(* IEC 61131-3 sources: stf-hw/web/public/sil, 1 file *)

(* ---- stf_plc.st ---- *)
(* STF Upgrade 12 - PLC program, IEC 61131-3 Structured Text. Generated by stf-cad/hbw/sil/iec.py *)
(* from the proven models; compile with MatIEC (iec2c). Task: 5 ms. *)

(* -1 / 0 / +1: which way to drive an axis toward its target; 0 inside the brake lead *)
FUNCTION Drive : INT
VAR_INPUT
    Pos, Tgt, Lead : REAL;
END_VAR
IF Tgt - Pos > Lead THEN Drive := 1; ELSIF Pos - Tgt > Lead THEN Drive := -1; ELSE Drive := 0; END_IF;
END_FUNCTION

(* HBW crane: travel, lift, Ausleger. Generated by stf-cad/hbw/sil/iec.py from the proven motion (control.py); do not edit. *)
FUNCTION_BLOCK FB_Crane
VAR_INPUT
    Enable : BOOL;        (* K0 safety relay OK AND mode = AUTO *)
    Ack : BOOL;           (* HMI acknowledge *)
    Reset : BOOL;         (* S3 reset, via the safety relay *)
    Cmd : INT;            (* job to start (0 = none), taken when READY *)
    Arg1 : INT;           (* binding: slot / bay / slot pair index *)
    I1 : BOOL;           (* reference switch horizontal *)
    I4 : BOOL;           (* reference switch vertical *)
    I5 : BOOL;           (* reference switch cantilever front *)
    I6 : BOOL;           (* reference switch cantilever back *)
    PosTravel : REAL;     (* travel, from the encoder counter *)
    PosLift : REAL;     (* lift, from the encoder counter *)
END_VAR
VAR_OUTPUT
    Q3 : BOOL;           (* horizontal towards rack (M2) *)
    Q4 : BOOL;           (* horizontal towards belt (M2) *)
    Q5 : BOOL;           (* vertical axis down (M3) *)
    Q6 : BOOL;           (* vertical axis up (M3) *)
    Q7 : BOOL;           (* cantilever forward (M4) *)
    Q8 : BOOL;           (* cantilever back (M4) *)
    Ready, Busy, Done, Fault : BOOL;   (* Done: one scan, when a job ends *)
    Alarm : INT;          (* the state whose watchdog tripped *)
    Sn : INT;             (* the active state *)
END_VAR
VAR
    Prev : INT := -1;
    Job, B1 : INT;
    Wd : TON;             (* step watchdog *)
    Tm : TON;             (* step timer *)
    WdTime : TIME;        (* the active state's watchdog; 0 = none *)
END_VAR
VAR CONSTANT
    TG_STORE_RETRIEVE_TRAVEL : ARRAY[1..143, 1..23] OF REAL := [0.0, 0.0, 0.0, 0.0, 0.0, 0.0, 0.0, 0.0, 0.0, 0.0, 0.0, 0.0, 0.0, 0.0, 0.0, 0.0, 0.0, 0.0, 0.0, 0.0, 0.0, 0.0, 0.0, 0.0, 0.0, 0.0, 0.0, 0.0, 120.0, 0.0, 0.0, 0.0, 0.0, 0.0, 240.0, 0.0, 0.0, 0.0, 0.0, 0.0, 665.0, 0.0, 0.0, 0.0, 0.0, 0.0, 0.0, 0.0, 0.0, 0.0, 0.0, 120.0, 0.0, 0.0, 0.0, 0.0, 0.0, 360.0, 0.0, 0.0, 0.0, 0.0, 0.0, 665.0, 0.0, 0.0, 0.0, 0.0, 0.0, 0.0, 0.0, 0.0, 0.0, 0.0, 120.0, 0.0, 0.0, 0.0, 0.0, 0.0, 480.0, 0.0, 0.0, 0.0, 0.0, 0.0, 665.0, 0.0, 0.0, 0.0, 0.0, 0.0, 0.0, 0.0, 0.0, 0.0, 0.0, 120.0, 0.0, 0.0, 0.0, 0.0, 0.0, 120.0, 0.0, 0.0, 0.0, 0.0, 0.0, 665.0, 0.0, 0.0, 0.0, 0.0, 0.0, 0.0, 0.0, 0.0, 0.0, 0.0, 120.0, 0.0, 0.0, 0.0, 0.0, 0.0, 240.0, 0.0, 0.0, 0.0, 0.0, 0.0, 665.0, 0.0, 0.0, 0.0, 0.0, 0.0, 0.0, 0.0, 0.0, 0.0, 0.0, 120.0, 0.0, 0.0, 0.0, 0.0, 0.0, 360.0, 0.0, 0.0, 0.0, 0.0, 0.0, 665.0, 0.0, 0.0, 0.0, 0.0, 0.0, 0.0, 0.0, 0.0, 0.0, 0.0, 120.0, 0.0, 0.0, 0.0, 0.0, 0.0, 480.0, 0.0, 0.0, 0.0, 0.0, 0.0, 665.0, 0.0, 0.0, 0.0, 0.0, 0.0, 0.0, 0.0, 0.0, 0.0, 0.0, 120.0, 0.0, 0.0, 0.0, 0.0, 0.0, 120.0, 0.0, 0.0, 0.0, 0.0, 0.0, 665.0, 0.0, 0.0, 0.0, 0.0, 0.0, 0.0, 0.0, 0.0, 0.0, 0.0, 120.0, 0.0, 0.0, 0.0, 0.0, 0.0, 240.0, 0.0, 0.0, 0.0, 0.0, 0.0, 665.0, 0.0, 0.0, 0.0, 0.0, 0.0, 0.0, 0.0, 0.0, 0.0, 0.0, 120.0, 0.0, 0.0, 0.0, 0.0, 0.0, 360.0, 0.0, 0.0, 0.0, 0.0, 0.0, 665.0, 0.0, 0.0, 0.0, 0.0, 0.0, 0.0, 0.0, 0.0, 0.0, 0.0, 120.0, 0.0, 0.0, 0.0, 0.0, 0.0, 480.0, 0.0, 0.0, 0.0, 0.0, 0.0, 665.0, 0.0, 0.0, 0.0, 0.0, 0.0, 0.0, 0.0, 0.0, 0.0, 0.0, 240.0, 0.0, 0.0, 0.0, 0.0, 0.0, 120.0, 0.0, 0.0, 0.0, 0.0, 0.0, 665.0, 0.0, 0.0, 0.0, 0.0, 0.0, 0.0, 0.0, 0.0, 0.0, 0.0, 0.0, 0.0, 0.0, 0.0, 0.0, 0.0, 0.0, 0.0, 0.0, 0.0, 0.0, 0.0, 0.0, 0.0, 0.0, 0.0, 0.0, 0.0, 0.0, 0.0, 0.0, 0.0, 0.0, 240.0, 0.0, 0.0, 0.0, 0.0, 0.0, 360.0, 0.0, 0.0, 0.0, 0.0, 0.0, 665.0, 0.0, 0.0, 0.0, 0.0, 0.0, 0.0, 0.0, 0.0, 0.0, 0.0, 240.0, 0.0, 0.0, 0.0, 0.0, 0.0, 480.0, 0.0, 0.0, 0.0, 0.0, 0.0, 665.0, 0.0, 0.0, 0.0, 0.0, 0.0, 0.0, 0.0, 0.0, 0.0, 0.0, 240.0, 0.0, 0.0, 0.0, 0.0, 0.0, 120.0, 0.0, 0.0, 0.0, 0.0, 0.0, 665.0, 0.0, 0.0, 0.0, 0.0, 0.0, 0.0, 0.0, 0.0, 0.0, 0.0, 240.0, 0.0, 0.0, 0.0, 0.0, 0.0, 240.0, 0.0, 0.0, 0.0, 0.0, 0.0, 665.0, 0.0, 0.0, 0.0, 0.0, 0.0, 0.0, 0.0, 0.0, 0.0, 0.0, 240.0, 0.0, 0.0, 0.0, 0.0, 0.0, 360.0, 0.0, 0.0, 0.0, 0.0, 0.0, 665.0, 0.0, 0.0, 0.0, 0.0, 0.0, 0.0, 0.0, 0.0, 0.0, 0.0, 240.0, 0.0, 0.0, 0.0, 0.0, 0.0, 480.0, 0.0, 0.0, 0.0, 0.0, 0.0, 665.0, 0.0, 0.0, 0.0, 0.0, 0.0, 0.0, 0.0, 0.0, 0.0, 0.0, 240.0, 0.0, 0.0, 0.0, 0.0, 0.0, 120.0, 0.0, 0.0, 0.0, 0.0, 0.0, 665.0, 0.0, 0.0, 0.0, 0.0, 0.0, 0.0, 0.0, 0.0, 0.0, 0.0, 240.0, 0.0, 0.0, 0.0, 0.0, 0.0, 240.0, 0.0, 0.0, 0.0, 0.0, 0.0, 665.0, 0.0, 0.0, 0.0, 0.0, 0.0, 0.0, 0.0, 0.0, 0.0, 0.0, 240.0, 0.0, 0.0, 0.0, 0.0, 0.0, 360.0, 0.0, 0.0, 0.0, 0.0, 0.0, 665.0, 0.0, 0.0, 0.0, 0.0, 0.0, 0.0, 0.0, 0.0, 0.0, 0.0, 240.0, 0.0, 0.0, 0.0, 0.0, 0.0, 480.0, 0.0, 0.0, 0.0, 0.0, 0.0, 665.0, 0.0, 0.0, 0.0, 0.0, 0.0, 0.0, 0.0, 0.0, 0.0, 0.0, 360.0, 0.0, 0.0, 0.0, 0.0, 0.0, 120.0, 0.0, 0.0, 0.0, 0.0, 0.0, 665.0, 0.0, 0.0, 0.0, 0.0, 0.0, 0.0, 0.0, 0.0, 0.0, 0.0, 360.0, 0.0, 0.0, 0.0, 0.0, 0.0, 240.0, 0.0, 0.0, 0.0, 0.0, 0.0, 665.0, 0.0, 0.0, 0.0, 0.0, 0.0, 0.0, 0.0, 0.0, 0.0, 0.0, 0.0, 0.0, 0.0, 0.0, 0.0, 0.0, 0.0, 0.0, 0.0, 0.0, 0.0, 0.0, 0.0, 0.0, 0.0, 0.0, 0.0, 0.0, 0.0, 0.0, 0.0, 0.0, 0.0, 360.0, 0.0, 0.0, 0.0, 0.0, 0.0, 480.0, 0.0, 0.0, 0.0, 0.0, 0.0, 665.0, 0.0, 0.0, 0.0, 0.0, 0.0, 0.0, 0.0, 0.0, 0.0, 0.0, 360.0, 0.0, 0.0, 0.0, 0.0, 0.0, 120.0, 0.0, 0.0, 0.0, 0.0, 0.0, 665.0, 0.0, 0.0, 0.0, 0.0, 0.0, 0.0, 0.0, 0.0, 0.0, 0.0, 360.0, 0.0, 0.0, 0.0, 0.0, 0.0, 240.0, 0.0, 0.0, 0.0, 0.0, 0.0, 665.0, 0.0, 0.0, 0.0, 0.0, 0.0, 0.0, 0.0, 0.0, 0.0, 0.0, 360.0, 0.0, 0.0, 0.0, 0.0, 0.0, 360.0, 0.0, 0.0, 0.0, 0.0, 0.0, 665.0, 0.0, 0.0, 0.0, 0.0, 0.0, 0.0, 0.0, 0.0, 0.0, 0.0, 360.0, 0.0, 0.0, 0.0, 0.0, 0.0, 480.0, 0.0, 0.0, 0.0, 0.0, 0.0, 665.0, 0.0, 0.0, 0.0, 0.0, 0.0, 0.0, 0.0, 0.0, 0.0, 0.0, 360.0, 0.0, 0.0, 0.0, 0.0, 0.0, 120.0, 0.0, 0.0, 0.0, 0.0, 0.0, 665.0, 0.0, 0.0, 0.0, 0.0, 0.0, 0.0, 0.0, 0.0, 0.0, 0.0, 360.0, 0.0, 0.0, 0.0, 0.0, 0.0, 240.0, 0.0, 0.0, 0.0, 0.0, 0.0, 665.0, 0.0, 0.0, 0.0, 0.0, 0.0, 0.0, 0.0, 0.0, 0.0, 0.0, 360.0, 0.0, 0.0, 0.0, 0.0, 0.0, 360.0, 0.0, 0.0, 0.0, 0.0, 0.0, 665.0, 0.0, 0.0, 0.0, 0.0, 0.0, 0.0, 0.0, 0.0, 0.0, 0.0, 360.0, 0.0, 0.0, 0.0, 0.0, 0.0, 480.0, 0.0, 0.0, 0.0, 0.0, 0.0, 665.0, 0.0, 0.0, 0.0, 0.0, 0.0, 0.0, 0.0, 0.0, 0.0, 0.0, 480.0, 0.0, 0.0, 0.0, 0.0, 0.0, 120.0, 0.0, 0.0, 0.0, 0.0, 0.0, 665.0, 0.0, 0.0, 0.0, 0.0, 0.0, 0.0, 0.0, 0.0, 0.0, 0.0, 480.0, 0.0, 0.0, 0.0, 0.0, 0.0, 240.0, 0.0, 0.0, 0.0, 0.0, 0.0, 665.0, 0.0, 0.0, 0.0, 0.0, 0.0, 0.0, 0.0, 0.0, 0.0, 0.0, 480.0, 0.0, 0.0, 0.0, 0.0, 0.0, 360.0, 0.0, 0.0, 0.0, 0.0, 0.0, 665.0, 0.0, 0.0, 0.0, 0.0, 0.0, 0.0, 0.0, 0.0, 0.0, 0.0, 0.0, 0.0, 0.0, 0.0, 0.0, 0.0, 0.0, 0.0, 0.0, 0.0, 0.0, 0.0, 0.0, 0.0, 0.0, 0.0, 0.0, 0.0, 0.0, 0.0, 0.0, 0.0, 0.0, 480.0, 0.0, 0.0, 0.0, 0.0, 0.0, 120.0, 0.0, 0.0, 0.0, 0.0, 0.0, 665.0, 0.0, 0.0, 0.0, 0.0, 0.0, 0.0, 0.0, 0.0, 0.0, 0.0, 480.0, 0.0, 0.0, 0.0, 0.0, 0.0, 240.0, 0.0, 0.0, 0.0, 0.0, 0.0, 665.0, 0.0, 0.0, 0.0, 0.0, 0.0, 0.0, 0.0, 0.0, 0.0, 0.0, 480.0, 0.0, 0.0, 0.0, 0.0, 0.0, 360.0, 0.0, 0.0, 0.0, 0.0, 0.0, 665.0, 0.0, 0.0, 0.0, 0.0, 0.0, 0.0, 0.0, 0.0, 0.0, 0.0, 480.0, 0.0, 0.0, 0.0, 0.0, 0.0, 480.0, 0.0, 0.0, 0.0, 0.0, 0.0, 665.0, 0.0, 0.0, 0.0, 0.0, 0.0, 0.0, 0.0, 0.0, 0.0, 0.0, 480.0, 0.0, 0.0, 0.0, 0.0, 0.0, 120.0, 0.0, 0.0, 0.0, 0.0, 0.0, 665.0, 0.0, 0.0, 0.0, 0.0, 0.0, 0.0, 0.0, 0.0, 0.0, 0.0, 480.0, 0.0, 0.0, 0.0, 0.0, 0.0, 240.0, 0.0, 0.0, 0.0, 0.0, 0.0, 665.0, 0.0, 0.0, 0.0, 0.0, 0.0, 0.0, 0.0, 0.0, 0.0, 0.0, 480.0, 0.0, 0.0, 0.0, 0.0, 0.0, 360.0, 0.0, 0.0, 0.0, 0.0, 0.0, 665.0, 0.0, 0.0, 0.0, 0.0, 0.0, 0.0, 0.0, 0.0, 0.0, 0.0, 480.0, 0.0, 0.0, 0.0, 0.0, 0.0, 480.0, 0.0, 0.0, 0.0, 0.0, 0.0, 665.0, 0.0, 0.0, 0.0, 0.0, 0.0, 0.0, 0.0, 0.0, 0.0, 0.0, 120.0, 0.0, 0.0, 0.0, 0.0, 0.0, 120.0, 0.0, 0.0, 0.0, 0.0, 0.0, 665.0, 0.0, 0.0, 0.0, 0.0, 0.0, 0.0, 0.0, 0.0, 0.0, 0.0, 120.0, 0.0, 0.0, 0.0, 0.0, 0.0, 240.0, 0.0, 0.0, 0.0, 0.0, 0.0, 665.0, 0.0, 0.0, 0.0, 0.0, 0.0, 0.0, 0.0, 0.0, 0.0, 0.0, 120.0, 0.0, 0.0, 0.0, 0.0, 0.0, 360.0, 0.0, 0.0, 0.0, 0.0, 0.0, 665.0, 0.0, 0.0, 0.0, 0.0, 0.0, 0.0, 0.0, 0.0, 0.0, 0.0, 120.0, 0.0, 0.0, 0.0, 0.0, 0.0, 480.0, 0.0, 0.0, 0.0, 0.0, 0.0, 665.0, 0.0, 0.0, 0.0, 0.0, 0.0, 0.0, 0.0, 0.0, 0.0, 0.0, 0.0, 0.0, 0.0, 0.0, 0.0, 0.0, 0.0, 0.0, 0.0, 0.0, 0.0, 0.0, 0.0, 0.0, 0.0, 0.0, 0.0, 0.0, 0.0, 0.0, 0.0, 0.0, 0.0, 120.0, 0.0, 0.0, 0.0, 0.0, 0.0, 240.0, 0.0, 0.0, 0.0, 0.0, 0.0, 665.0, 0.0, 0.0, 0.0, 0.0, 0.0, 0.0, 0.0, 0.0, 0.0, 0.0, 120.0, 0.0, 0.0, 0.0, 0.0, 0.0, 360.0, 0.0, 0.0, 0.0, 0.0, 0.0, 665.0, 0.0, 0.0, 0.0, 0.0, 0.0, 0.0, 0.0, 0.0, 0.0, 0.0, 120.0, 0.0, 0.0, 0.0, 0.0, 0.0, 480.0, 0.0, 0.0, 0.0, 0.0, 0.0, 665.0, 0.0, 0.0, 0.0, 0.0, 0.0, 0.0, 0.0, 0.0, 0.0, 0.0, 120.0, 0.0, 0.0, 0.0, 0.0, 0.0, 120.0, 0.0, 0.0, 0.0, 0.0, 0.0, 665.0, 0.0, 0.0, 0.0, 0.0, 0.0, 0.0, 0.0, 0.0, 0.0, 0.0, 120.0, 0.0, 0.0, 0.0, 0.0, 0.0, 240.0, 0.0, 0.0, 0.0, 0.0, 0.0, 665.0, 0.0, 0.0, 0.0, 0.0, 0.0, 0.0, 0.0, 0.0, 0.0, 0.0, 120.0, 0.0, 0.0, 0.0, 0.0, 0.0, 360.0, 0.0, 0.0, 0.0, 0.0, 0.0, 665.0, 0.0, 0.0, 0.0, 0.0, 0.0, 0.0, 0.0, 0.0, 0.0, 0.0, 120.0, 0.0, 0.0, 0.0, 0.0, 0.0, 480.0, 0.0, 0.0, 0.0, 0.0, 0.0, 665.0, 0.0, 0.0, 0.0, 0.0, 0.0, 0.0, 0.0, 0.0, 0.0, 0.0, 240.0, 0.0, 0.0, 0.0, 0.0, 0.0, 120.0, 0.0, 0.0, 0.0, 0.0, 0.0, 665.0, 0.0, 0.0, 0.0, 0.0, 0.0, 0.0, 0.0, 0.0, 0.0, 0.0, 240.0, 0.0, 0.0, 0.0, 0.0, 0.0, 240.0, 0.0, 0.0, 0.0, 0.0, 0.0, 665.0, 0.0, 0.0, 0.0, 0.0, 0.0, 0.0, 0.0, 0.0, 0.0, 0.0, 240.0, 0.0, 0.0, 0.0, 0.0, 0.0, 360.0, 0.0, 0.0, 0.0, 0.0, 0.0, 665.0, 0.0, 0.0, 0.0, 0.0, 0.0, 0.0, 0.0, 0.0, 0.0, 0.0, 240.0, 0.0, 0.0, 0.0, 0.0, 0.0, 480.0, 0.0, 0.0, 0.0, 0.0, 0.0, 665.0, 0.0, 0.0, 0.0, 0.0, 0.0, 0.0, 0.0, 0.0, 0.0, 0.0, 240.0, 0.0, 0.0, 0.0, 0.0, 0.0, 120.0, 0.0, 0.0, 0.0, 0.0, 0.0, 665.0, 0.0, 0.0, 0.0, 0.0, 0.0, 0.0, 0.0, 0.0, 0.0, 0.0, 0.0, 0.0, 0.0, 0.0, 0.0, 0.0, 0.0, 0.0, 0.0, 0.0, 0.0, 0.0, 0.0, 0.0, 0.0, 0.0, 0.0, 0.0, 0.0, 0.0, 0.0, 0.0, 0.0, 240.0, 0.0, 0.0, 0.0, 0.0, 0.0, 360.0, 0.0, 0.0, 0.0, 0.0, 0.0, 665.0, 0.0, 0.0, 0.0, 0.0, 0.0, 0.0, 0.0, 0.0, 0.0, 0.0, 240.0, 0.0, 0.0, 0.0, 0.0, 0.0, 480.0, 0.0, 0.0, 0.0, 0.0, 0.0, 665.0, 0.0, 0.0, 0.0, 0.0, 0.0, 0.0, 0.0, 0.0, 0.0, 0.0, 240.0, 0.0, 0.0, 0.0, 0.0, 0.0, 120.0, 0.0, 0.0, 0.0, 0.0, 0.0, 665.0, 0.0, 0.0, 0.0, 0.0, 0.0, 0.0, 0.0, 0.0, 0.0, 0.0, 240.0, 0.0, 0.0, 0.0, 0.0, 0.0, 240.0, 0.0, 0.0, 0.0, 0.0, 0.0, 665.0, 0.0, 0.0, 0.0, 0.0, 0.0, 0.0, 0.0, 0.0, 0.0, 0.0, 240.0, 0.0, 0.0, 0.0, 0.0, 0.0, 360.0, 0.0, 0.0, 0.0, 0.0, 0.0, 665.0, 0.0, 0.0, 0.0, 0.0, 0.0, 0.0, 0.0, 0.0, 0.0, 0.0, 240.0, 0.0, 0.0, 0.0, 0.0, 0.0, 480.0, 0.0, 0.0, 0.0, 0.0, 0.0, 665.0, 0.0, 0.0, 0.0, 0.0, 0.0, 0.0, 0.0, 0.0, 0.0, 0.0, 360.0, 0.0, 0.0, 0.0, 0.0, 0.0, 120.0, 0.0, 0.0, 0.0, 0.0, 0.0, 665.0, 0.0, 0.0, 0.0, 0.0, 0.0, 0.0, 0.0, 0.0, 0.0, 0.0, 360.0, 0.0, 0.0, 0.0, 0.0, 0.0, 240.0, 0.0, 0.0, 0.0, 0.0, 0.0, 665.0, 0.0, 0.0, 0.0, 0.0, 0.0, 0.0, 0.0, 0.0, 0.0, 0.0, 360.0, 0.0, 0.0, 0.0, 0.0, 0.0, 360.0, 0.0, 0.0, 0.0, 0.0, 0.0, 665.0, 0.0, 0.0, 0.0, 0.0, 0.0, 0.0, 0.0, 0.0, 0.0, 0.0, 360.0, 0.0, 0.0, 0.0, 0.0, 0.0, 480.0, 0.0, 0.0, 0.0, 0.0, 0.0, 665.0, 0.0, 0.0, 0.0, 0.0, 0.0, 0.0, 0.0, 0.0, 0.0, 0.0, 360.0, 0.0, 0.0, 0.0, 0.0, 0.0, 120.0, 0.0, 0.0, 0.0, 0.0, 0.0, 665.0, 0.0, 0.0, 0.0, 0.0, 0.0, 0.0, 0.0, 0.0, 0.0, 0.0, 360.0, 0.0, 0.0, 0.0, 0.0, 0.0, 240.0, 0.0, 0.0, 0.0, 0.0, 0.0, 665.0, 0.0, 0.0, 0.0, 0.0, 0.0, 0.0, 0.0, 0.0, 0.0, 0.0, 0.0, 0.0, 0.0, 0.0, 0.0, 0.0, 0.0, 0.0, 0.0, 0.0, 0.0, 0.0, 0.0, 0.0, 0.0, 0.0, 0.0, 0.0, 0.0, 0.0, 0.0, 0.0, 0.0, 360.0, 0.0, 0.0, 0.0, 0.0, 0.0, 480.0, 0.0, 0.0, 0.0, 0.0, 0.0, 665.0, 0.0, 0.0, 0.0, 0.0, 0.0, 0.0, 0.0, 0.0, 0.0, 0.0, 360.0, 0.0, 0.0, 0.0, 0.0, 0.0, 120.0, 0.0, 0.0, 0.0, 0.0, 0.0, 665.0, 0.0, 0.0, 0.0, 0.0, 0.0, 0.0, 0.0, 0.0, 0.0, 0.0, 360.0, 0.0, 0.0, 0.0, 0.0, 0.0, 240.0, 0.0, 0.0, 0.0, 0.0, 0.0, 665.0, 0.0, 0.0, 0.0, 0.0, 0.0, 0.0, 0.0, 0.0, 0.0, 0.0, 360.0, 0.0, 0.0, 0.0, 0.0, 0.0, 360.0, 0.0, 0.0, 0.0, 0.0, 0.0, 665.0, 0.0, 0.0, 0.0, 0.0, 0.0, 0.0, 0.0, 0.0, 0.0, 0.0, 360.0, 0.0, 0.0, 0.0, 0.0, 0.0, 480.0, 0.0, 0.0, 0.0, 0.0, 0.0, 665.0, 0.0, 0.0, 0.0, 0.0, 0.0, 0.0, 0.0, 0.0, 0.0, 0.0, 480.0, 0.0, 0.0, 0.0, 0.0, 0.0, 120.0, 0.0, 0.0, 0.0, 0.0, 0.0, 665.0, 0.0, 0.0, 0.0, 0.0, 0.0, 0.0, 0.0, 0.0, 0.0, 0.0, 480.0, 0.0, 0.0, 0.0, 0.0, 0.0, 240.0, 0.0, 0.0, 0.0, 0.0, 0.0, 665.0, 0.0, 0.0, 0.0, 0.0, 0.0, 0.0, 0.0, 0.0, 0.0, 0.0, 480.0, 0.0, 0.0, 0.0, 0.0, 0.0, 360.0, 0.0, 0.0, 0.0, 0.0, 0.0, 665.0, 0.0, 0.0, 0.0, 0.0, 0.0, 0.0, 0.0, 0.0, 0.0, 0.0, 480.0, 0.0, 0.0, 0.0, 0.0, 0.0, 480.0, 0.0, 0.0, 0.0, 0.0, 0.0, 665.0, 0.0, 0.0, 0.0, 0.0, 0.0, 0.0, 0.0, 0.0, 0.0, 0.0, 480.0, 0.0, 0.0, 0.0, 0.0, 0.0, 120.0, 0.0, 0.0, 0.0, 0.0, 0.0, 665.0, 0.0, 0.0, 0.0, 0.0, 0.0, 0.0, 0.0, 0.0, 0.0, 0.0, 480.0, 0.0, 0.0, 0.0, 0.0, 0.0, 240.0, 0.0, 0.0, 0.0, 0.0, 0.0, 665.0, 0.0, 0.0, 0.0, 0.0, 0.0, 0.0, 0.0, 0.0, 0.0, 0.0, 480.0, 0.0, 0.0, 0.0, 0.0, 0.0, 360.0, 0.0, 0.0, 0.0, 0.0, 0.0, 665.0, 0.0, 0.0, 0.0, 0.0, 0.0, 0.0, 0.0, 0.0, 0.0, 0.0, 0.0, 0.0, 0.0, 0.0, 0.0, 0.0, 0.0, 0.0, 0.0, 0.0, 0.0, 0.0, 0.0, 0.0, 0.0, 0.0, 0.0, 0.0, 0.0, 0.0, 0.0, 0.0, 0.0, 480.0, 0.0, 0.0, 0.0, 0.0, 0.0, 120.0, 0.0, 0.0, 0.0, 0.0, 0.0, 665.0, 0.0, 0.0, 0.0, 0.0, 0.0, 0.0, 0.0, 0.0, 0.0, 0.0, 480.0, 0.0, 0.0, 0.0, 0.0, 0.0, 240.0, 0.0, 0.0, 0.0, 0.0, 0.0, 665.0, 0.0, 0.0, 0.0, 0.0, 0.0, 0.0, 0.0, 0.0, 0.0, 0.0, 480.0, 0.0, 0.0, 0.0, 0.0, 0.0, 360.0, 0.0, 0.0, 0.0, 0.0, 0.0, 665.0, 0.0, 0.0, 0.0, 0.0, 0.0, 0.0, 0.0, 0.0, 0.0, 0.0, 480.0, 0.0, 0.0, 0.0, 0.0, 0.0, 480.0, 0.0, 0.0, 0.0, 0.0, 0.0, 665.0, 0.0, 0.0, 0.0, 0.0, 0.0, 0.0, 0.0, 0.0, 0.0, 0.0, 120.0, 0.0, 0.0, 0.0, 0.0, 0.0, 120.0, 0.0, 0.0, 0.0, 0.0, 0.0, 665.0, 0.0, 0.0, 0.0, 0.0, 0.0, 0.0, 0.0, 0.0, 0.0, 0.0, 120.0, 0.0, 0.0, 0.0, 0.0, 0.0, 240.0, 0.0, 0.0, 0.0, 0.0, 0.0, 665.0, 0.0, 0.0, 0.0, 0.0, 0.0, 0.0, 0.0, 0.0, 0.0, 0.0, 120.0, 0.0, 0.0, 0.0, 0.0, 0.0, 360.0, 0.0, 0.0, 0.0, 0.0, 0.0, 665.0, 0.0, 0.0, 0.0, 0.0, 0.0, 0.0, 0.0, 0.0, 0.0, 0.0, 120.0, 0.0, 0.0, 0.0, 0.0, 0.0, 480.0, 0.0, 0.0, 0.0, 0.0, 0.0, 665.0, 0.0, 0.0, 0.0, 0.0, 0.0, 0.0, 0.0, 0.0, 0.0, 0.0, 120.0, 0.0, 0.0, 0.0, 0.0, 0.0, 120.0, 0.0, 0.0, 0.0, 0.0, 0.0, 665.0, 0.0, 0.0, 0.0, 0.0, 0.0, 0.0, 0.0, 0.0, 0.0, 0.0, 120.0, 0.0, 0.0, 0.0, 0.0, 0.0, 240.0, 0.0, 0.0, 0.0, 0.0, 0.0, 665.0, 0.0, 0.0, 0.0, 0.0, 0.0, 0.0, 0.0, 0.0, 0.0, 0.0, 120.0, 0.0, 0.0, 0.0, 0.0, 0.0, 360.0, 0.0, 0.0, 0.0, 0.0, 0.0, 665.0, 0.0, 0.0, 0.0, 0.0, 0.0, 0.0, 0.0, 0.0, 0.0, 0.0, 120.0, 0.0, 0.0, 0.0, 0.0, 0.0, 480.0, 0.0, 0.0, 0.0, 0.0, 0.0, 665.0, 0.0, 0.0, 0.0, 0.0, 0.0, 0.0, 0.0, 0.0, 0.0, 0.0, 0.0, 0.0, 0.0, 0.0, 0.0, 0.0, 0.0, 0.0, 0.0, 0.0, 0.0, 0.0, 0.0, 0.0, 0.0, 0.0, 0.0, 0.0, 0.0, 0.0, 0.0, 0.0, 0.0, 120.0, 0.0, 0.0, 0.0, 0.0, 0.0, 240.0, 0.0, 0.0, 0.0, 0.0, 0.0, 665.0, 0.0, 0.0, 0.0, 0.0, 0.0, 0.0, 0.0, 0.0, 0.0, 0.0, 120.0, 0.0, 0.0, 0.0, 0.0, 0.0, 360.0, 0.0, 0.0, 0.0, 0.0, 0.0, 665.0, 0.0, 0.0, 0.0, 0.0, 0.0, 0.0, 0.0, 0.0, 0.0, 0.0, 120.0, 0.0, 0.0, 0.0, 0.0, 0.0, 480.0, 0.0, 0.0, 0.0, 0.0, 0.0, 665.0, 0.0, 0.0, 0.0, 0.0, 0.0, 0.0, 0.0, 0.0, 0.0, 0.0, 240.0, 0.0, 0.0, 0.0, 0.0, 0.0, 120.0, 0.0, 0.0, 0.0, 0.0, 0.0, 665.0, 0.0, 0.0, 0.0, 0.0, 0.0, 0.0, 0.0, 0.0, 0.0, 0.0, 240.0, 0.0, 0.0, 0.0, 0.0, 0.0, 240.0, 0.0, 0.0, 0.0, 0.0, 0.0, 665.0, 0.0, 0.0, 0.0, 0.0, 0.0, 0.0, 0.0, 0.0, 0.0, 0.0, 240.0, 0.0, 0.0, 0.0, 0.0, 0.0, 360.0, 0.0, 0.0, 0.0, 0.0, 0.0, 665.0, 0.0, 0.0, 0.0, 0.0, 0.0, 0.0, 0.0, 0.0, 0.0, 0.0, 240.0, 0.0, 0.0, 0.0, 0.0, 0.0, 480.0, 0.0, 0.0, 0.0, 0.0, 0.0, 665.0, 0.0, 0.0, 0.0, 0.0, 0.0, 0.0, 0.0, 0.0, 0.0, 0.0, 240.0, 0.0, 0.0, 0.0, 0.0, 0.0, 120.0, 0.0, 0.0, 0.0, 0.0, 0.0, 665.0, 0.0, 0.0, 0.0, 0.0, 0.0, 0.0, 0.0, 0.0, 0.0, 0.0, 240.0, 0.0, 0.0, 0.0, 0.0, 0.0, 240.0, 0.0, 0.0, 0.0, 0.0, 0.0, 665.0, 0.0, 0.0, 0.0, 0.0, 0.0, 0.0, 0.0, 0.0, 0.0, 0.0, 240.0, 0.0, 0.0, 0.0, 0.0, 0.0, 360.0, 0.0, 0.0, 0.0, 0.0, 0.0, 665.0, 0.0, 0.0, 0.0, 0.0, 0.0, 0.0, 0.0, 0.0, 0.0, 0.0, 240.0, 0.0, 0.0, 0.0, 0.0, 0.0, 480.0, 0.0, 0.0, 0.0, 0.0, 0.0, 665.0, 0.0, 0.0, 0.0, 0.0, 0.0, 0.0, 0.0, 0.0, 0.0, 0.0, 240.0, 0.0, 0.0, 0.0, 0.0, 0.0, 120.0, 0.0, 0.0, 0.0, 0.0, 0.0, 665.0, 0.0, 0.0, 0.0, 0.0, 0.0, 0.0, 0.0, 0.0, 0.0, 0.0, 0.0, 0.0, 0.0, 0.0, 0.0, 0.0, 0.0, 0.0, 0.0, 0.0, 0.0, 0.0, 0.0, 0.0, 0.0, 0.0, 0.0, 0.0, 0.0, 0.0, 0.0, 0.0, 0.0, 240.0, 0.0, 0.0, 0.0, 0.0, 0.0, 360.0, 0.0, 0.0, 0.0, 0.0, 0.0, 665.0, 0.0, 0.0, 0.0, 0.0, 0.0, 0.0, 0.0, 0.0, 0.0, 0.0, 240.0, 0.0, 0.0, 0.0, 0.0, 0.0, 480.0, 0.0, 0.0, 0.0, 0.0, 0.0, 665.0, 0.0, 0.0, 0.0, 0.0, 0.0, 0.0, 0.0, 0.0, 0.0, 0.0, 360.0, 0.0, 0.0, 0.0, 0.0, 0.0, 120.0, 0.0, 0.0, 0.0, 0.0, 0.0, 665.0, 0.0, 0.0, 0.0, 0.0, 0.0, 0.0, 0.0, 0.0, 0.0, 0.0, 360.0, 0.0, 0.0, 0.0, 0.0, 0.0, 240.0, 0.0, 0.0, 0.0, 0.0, 0.0, 665.0, 0.0, 0.0, 0.0, 0.0, 0.0, 0.0, 0.0, 0.0, 0.0, 0.0, 360.0, 0.0, 0.0, 0.0, 0.0, 0.0, 360.0, 0.0, 0.0, 0.0, 0.0, 0.0, 665.0, 0.0, 0.0, 0.0, 0.0, 0.0, 0.0, 0.0, 0.0, 0.0, 0.0, 360.0, 0.0, 0.0, 0.0, 0.0, 0.0, 480.0, 0.0, 0.0, 0.0, 0.0, 0.0, 665.0, 0.0, 0.0, 0.0, 0.0, 0.0, 0.0, 0.0, 0.0, 0.0, 0.0, 360.0, 0.0, 0.0, 0.0, 0.0, 0.0, 120.0, 0.0, 0.0, 0.0, 0.0, 0.0, 665.0, 0.0, 0.0, 0.0, 0.0, 0.0, 0.0, 0.0, 0.0, 0.0, 0.0, 360.0, 0.0, 0.0, 0.0, 0.0, 0.0, 240.0, 0.0, 0.0, 0.0, 0.0, 0.0, 665.0, 0.0, 0.0, 0.0, 0.0, 0.0, 0.0, 0.0, 0.0, 0.0, 0.0, 360.0, 0.0, 0.0, 0.0, 0.0, 0.0, 360.0, 0.0, 0.0, 0.0, 0.0, 0.0, 665.0, 0.0, 0.0, 0.0, 0.0, 0.0, 0.0, 0.0, 0.0, 0.0, 0.0, 360.0, 0.0, 0.0, 0.0, 0.0, 0.0, 480.0, 0.0, 0.0, 0.0, 0.0, 0.0, 665.0, 0.0, 0.0, 0.0, 0.0, 0.0, 0.0, 0.0, 0.0, 0.0, 0.0, 360.0, 0.0, 0.0, 0.0, 0.0, 0.0, 120.0, 0.0, 0.0, 0.0, 0.0, 0.0, 665.0, 0.0, 0.0, 0.0, 0.0, 0.0, 0.0, 0.0, 0.0, 0.0, 0.0, 360.0, 0.0, 0.0, 0.0, 0.0, 0.0, 240.0, 0.0, 0.0, 0.0, 0.0, 0.0, 665.0, 0.0, 0.0, 0.0, 0.0, 0.0, 0.0, 0.0, 0.0, 0.0, 0.0, 0.0, 0.0, 0.0, 0.0, 0.0, 0.0, 0.0, 0.0, 0.0, 0.0, 0.0, 0.0, 0.0, 0.0, 0.0, 0.0, 0.0, 0.0, 0.0, 0.0, 0.0, 0.0, 0.0, 360.0, 0.0, 0.0, 0.0, 0.0, 0.0, 480.0, 0.0, 0.0, 0.0, 0.0, 0.0, 665.0, 0.0, 0.0, 0.0, 0.0, 0.0, 0.0, 0.0, 0.0, 0.0, 0.0, 480.0, 0.0, 0.0, 0.0, 0.0, 0.0, 120.0, 0.0, 0.0, 0.0, 0.0, 0.0, 665.0, 0.0, 0.0, 0.0, 0.0, 0.0, 0.0, 0.0, 0.0, 0.0, 0.0, 480.0, 0.0, 0.0, 0.0, 0.0, 0.0, 240.0, 0.0, 0.0, 0.0, 0.0, 0.0, 665.0, 0.0, 0.0, 0.0, 0.0, 0.0, 0.0, 0.0, 0.0, 0.0, 0.0, 480.0, 0.0, 0.0, 0.0, 0.0, 0.0, 360.0, 0.0, 0.0, 0.0, 0.0, 0.0, 665.0, 0.0, 0.0, 0.0, 0.0, 0.0, 0.0, 0.0, 0.0, 0.0, 0.0, 480.0, 0.0, 0.0, 0.0, 0.0, 0.0, 480.0, 0.0, 0.0, 0.0, 0.0, 0.0, 665.0, 0.0, 0.0, 0.0, 0.0, 0.0, 0.0, 0.0, 0.0, 0.0, 0.0, 480.0, 0.0, 0.0, 0.0, 0.0, 0.0, 120.0, 0.0, 0.0, 0.0, 0.0, 0.0, 665.0, 0.0, 0.0, 0.0, 0.0, 0.0, 0.0, 0.0, 0.0, 0.0, 0.0, 480.0, 0.0, 0.0, 0.0, 0.0, 0.0, 240.0, 0.0, 0.0, 0.0, 0.0, 0.0, 665.0, 0.0, 0.0, 0.0, 0.0, 0.0, 0.0, 0.0, 0.0, 0.0, 0.0, 480.0, 0.0, 0.0, 0.0, 0.0, 0.0, 360.0, 0.0, 0.0, 0.0, 0.0, 0.0, 665.0, 0.0, 0.0, 0.0, 0.0, 0.0, 0.0, 0.0, 0.0, 0.0, 0.0, 480.0, 0.0, 0.0, 0.0, 0.0, 0.0, 480.0, 0.0, 0.0, 0.0, 0.0, 0.0, 665.0, 0.0, 0.0, 0.0, 0.0, 0.0, 0.0, 0.0, 0.0, 0.0, 0.0, 480.0, 0.0, 0.0, 0.0, 0.0, 0.0, 120.0, 0.0, 0.0, 0.0, 0.0, 0.0, 665.0, 0.0, 0.0, 0.0, 0.0, 0.0, 0.0, 0.0, 0.0, 0.0, 0.0, 480.0, 0.0, 0.0, 0.0, 0.0, 0.0, 240.0, 0.0, 0.0, 0.0, 0.0, 0.0, 665.0, 0.0, 0.0, 0.0, 0.0, 0.0, 0.0, 0.0, 0.0, 0.0, 0.0, 480.0, 0.0, 0.0, 0.0, 0.0, 0.0, 360.0, 0.0, 0.0, 0.0, 0.0, 0.0, 665.0, 0.0, 0.0, 0.0, 0.0, 0.0];
    TG_STORE_RETRIEVE_LIFT : ARRAY[1..143, 1..23] OF REAL := [0.0, 0.0, 0.0, 0.0, 0.0, 0.0, 0.0, 0.0, 0.0, 0.0, 0.0, 0.0, 0.0, 0.0, 0.0, 0.0, 0.0, 0.0, 0.0, 0.0, 0.0, 0.0, 0.0, 80.0, 0.0, 100.0, 0.0, 260.0, 0.0, 120.0, 0.0, 100.0, 0.0, 260.0, 0.0, 100.0, 0.0, 120.0, 0.0, 260.0, 0.0, 100.0, 0.0, 80.0, 0.0, 260.0, 80.0, 0.0, 100.0, 0.0, 260.0, 0.0, 120.0, 0.0, 100.0, 0.0, 260.0, 0.0, 100.0, 0.0, 120.0, 0.0, 260.0, 0.0, 100.0, 0.0, 80.0, 0.0, 260.0, 80.0, 0.0, 100.0, 0.0, 260.0, 0.0, 120.0, 0.0, 100.0, 0.0, 260.0, 0.0, 100.0, 0.0, 120.0, 0.0, 260.0, 0.0, 100.0, 0.0, 80.0, 0.0, 260.0, 80.0, 0.0, 100.0, 0.0, 260.0, 0.0, 120.0, 0.0, 100.0, 0.0, 260.0, 0.0, 220.0, 0.0, 240.0, 0.0, 260.0, 0.0, 100.0, 0.0, 80.0, 0.0, 260.0, 80.0, 0.0, 100.0, 0.0, 260.0, 0.0, 120.0, 0.0, 100.0, 0.0, 260.0, 0.0, 220.0, 0.0, 240.0, 0.0, 260.0, 0.0, 100.0, 0.0, 80.0, 0.0, 260.0, 80.0, 0.0, 100.0, 0.0, 260.0, 0.0, 120.0, 0.0, 100.0, 0.0, 260.0, 0.0, 220.0, 0.0, 240.0, 0.0, 260.0, 0.0, 100.0, 0.0, 80.0, 0.0, 260.0, 80.0, 0.0, 100.0, 0.0, 260.0, 0.0, 120.0, 0.0, 100.0, 0.0, 260.0, 0.0, 220.0, 0.0, 240.0, 0.0, 260.0, 0.0, 100.0, 0.0, 80.0, 0.0, 260.0, 80.0, 0.0, 100.0, 0.0, 260.0, 0.0, 120.0, 0.0, 100.0, 0.0, 260.0, 0.0, 340.0, 0.0, 360.0, 0.0, 260.0, 0.0, 100.0, 0.0, 80.0, 0.0, 260.0, 80.0, 0.0, 100.0, 0.0, 260.0, 0.0, 120.0, 0.0, 100.0, 0.0, 260.0, 0.0, 340.0, 0.0, 360.0, 0.0, 260.0, 0.0, 100.0, 0.0, 80.0, 0.0, 260.0, 80.0, 0.0, 100.0, 0.0, 260.0, 0.0, 120.0, 0.0, 100.0, 0.0, 260.0, 0.0, 340.0, 0.0, 360.0, 0.0, 260.0, 0.0, 100.0, 0.0, 80.0, 0.0, 260.0, 80.0, 0.0, 100.0, 0.0, 260.0, 0.0, 120.0, 0.0, 100.0, 0.0, 260.0, 0.0, 340.0, 0.0, 360.0, 0.0, 260.0, 0.0, 100.0, 0.0, 80.0, 0.0, 260.0, 80.0, 0.0, 100.0, 0.0, 260.0, 0.0, 120.0, 0.0, 100.0, 0.0, 260.0, 0.0, 100.0, 0.0, 120.0, 0.0, 260.0, 0.0, 100.0, 0.0, 80.0, 0.0, 260.0, 0.0, 0.0, 0.0, 0.0, 0.0, 0.0, 0.0, 0.0, 0.0, 0.0, 0.0, 0.0, 0.0, 0.0, 0.0, 0.0, 0.0, 0.0, 0.0, 0.0, 0.0, 0.0, 0.0, 80.0, 0.0, 100.0, 0.0, 260.0, 0.0, 120.0, 0.0, 100.0, 0.0, 260.0, 0.0, 100.0, 0.0, 120.0, 0.0, 260.0, 0.0, 100.0, 0.0, 80.0, 0.0, 260.0, 80.0, 0.0, 100.0, 0.0, 260.0, 0.0, 120.0, 0.0, 100.0, 0.0, 260.0, 0.0, 100.0, 0.0, 120.0, 0.0, 260.0, 0.0, 100.0, 0.0, 80.0, 0.0, 260.0, 80.0, 0.0, 100.0, 0.0, 260.0, 0.0, 120.0, 0.0, 100.0, 0.0, 260.0, 0.0, 220.0, 0.0, 240.0, 0.0, 260.0, 0.0, 100.0, 0.0, 80.0, 0.0, 260.0, 80.0, 0.0, 100.0, 0.0, 260.0, 0.0, 120.0, 0.0, 100.0, 0.0, 260.0, 0.0, 220.0, 0.0, 240.0, 0.0, 260.0, 0.0, 100.0, 0.0, 80.0, 0.0, 260.0, 80.0, 0.0, 100.0, 0.0, 260.0, 0.0, 120.0, 0.0, 100.0, 0.0, 260.0, 0.0, 220.0, 0.0, 240.0, 0.0, 260.0, 0.0, 100.0, 0.0, 80.0, 0.0, 260.0, 80.0, 0.0, 100.0, 0.0, 260.0, 0.0, 120.0, 0.0, 100.0, 0.0, 260.0, 0.0, 220.0, 0.0, 240.0, 0.0, 260.0, 0.0, 100.0, 0.0, 80.0, 0.0, 260.0, 80.0, 0.0, 100.0, 0.0, 260.0, 0.0, 120.0, 0.0, 100.0, 0.0, 260.0, 0.0, 340.0, 0.0, 360.0, 0.0, 260.0, 0.0, 100.0, 0.0, 80.0, 0.0, 260.0, 80.0, 0.0, 100.0, 0.0, 260.0, 0.0, 120.0, 0.0, 100.0, 0.0, 260.0, 0.0, 340.0, 0.0, 360.0, 0.0, 260.0, 0.0, 100.0, 0.0, 80.0, 0.0, 260.0, 80.0, 0.0, 100.0, 0.0, 260.0, 0.0, 120.0, 0.0, 100.0, 0.0, 260.0, 0.0, 340.0, 0.0, 360.0, 0.0, 260.0, 0.0, 100.0, 0.0, 80.0, 0.0, 260.0, 80.0, 0.0, 100.0, 0.0, 260.0, 0.0, 120.0, 0.0, 100.0, 0.0, 260.0, 0.0, 340.0, 0.0, 360.0, 0.0, 260.0, 0.0, 100.0, 0.0, 80.0, 0.0, 260.0, 80.0, 0.0, 100.0, 0.0, 260.0, 0.0, 120.0, 0.0, 100.0, 0.0, 260.0, 0.0, 100.0, 0.0, 120.0, 0.0, 260.0, 0.0, 100.0, 0.0, 80.0, 0.0, 260.0, 80.0, 0.0, 100.0, 0.0, 260.0, 0.0, 120.0, 0.0, 100.0, 0.0, 260.0, 0.0, 100.0, 0.0, 120.0, 0.0, 260.0, 0.0, 100.0, 0.0, 80.0, 0.0, 260.0, 0.0, 0.0, 0.0, 0.0, 0.0, 0.0, 0.0, 0.0, 0.0, 0.0, 0.0, 0.0, 0.0, 0.0, 0.0, 0.0, 0.0, 0.0, 0.0, 0.0, 0.0, 0.0, 0.0, 80.0, 0.0, 100.0, 0.0, 260.0, 0.0, 120.0, 0.0, 100.0, 0.0, 260.0, 0.0, 100.0, 0.0, 120.0, 0.0, 260.0, 0.0, 100.0, 0.0, 80.0, 0.0, 260.0, 80.0, 0.0, 100.0, 0.0, 260.0, 0.0, 120.0, 0.0, 100.0, 0.0, 260.0, 0.0, 220.0, 0.0, 240.0, 0.0, 260.0, 0.0, 100.0, 0.0, 80.0, 0.0, 260.0, 80.0, 0.0, 100.0, 0.0, 260.0, 0.0, 120.0, 0.0, 100.0, 0.0, 260.0, 0.0, 220.0, 0.0, 240.0, 0.0, 260.0, 0.0, 100.0, 0.0, 80.0, 0.0, 260.0, 80.0, 0.0, 100.0, 0.0, 260.0, 0.0, 120.0, 0.0, 100.0, 0.0, 260.0, 0.0, 220.0, 0.0, 240.0, 0.0, 260.0, 0.0, 100.0, 0.0, 80.0, 0.0, 260.0, 80.0, 0.0, 100.0, 0.0, 260.0, 0.0, 120.0, 0.0, 100.0, 0.0, 260.0, 0.0, 220.0, 0.0, 240.0, 0.0, 260.0, 0.0, 100.0, 0.0, 80.0, 0.0, 260.0, 80.0, 0.0, 100.0, 0.0, 260.0, 0.0, 120.0, 0.0, 100.0, 0.0, 260.0, 0.0, 340.0, 0.0, 360.0, 0.0, 260.0, 0.0, 100.0, 0.0, 80.0, 0.0, 260.0, 80.0, 0.0, 100.0, 0.0, 260.0, 0.0, 120.0, 0.0, 100.0, 0.0, 260.0, 0.0, 340.0, 0.0, 360.0, 0.0, 260.0, 0.0, 100.0, 0.0, 80.0, 0.0, 260.0, 80.0, 0.0, 100.0, 0.0, 260.0, 0.0, 120.0, 0.0, 100.0, 0.0, 260.0, 0.0, 340.0, 0.0, 360.0, 0.0, 260.0, 0.0, 100.0, 0.0, 80.0, 0.0, 260.0, 80.0, 0.0, 100.0, 0.0, 260.0, 0.0, 120.0, 0.0, 100.0, 0.0, 260.0, 0.0, 340.0, 0.0, 360.0, 0.0, 260.0, 0.0, 100.0, 0.0, 80.0, 0.0, 260.0, 80.0, 0.0, 100.0, 0.0, 260.0, 0.0, 120.0, 0.0, 100.0, 0.0, 260.0, 0.0, 100.0, 0.0, 120.0, 0.0, 260.0, 0.0, 100.0, 0.0, 80.0, 0.0, 260.0, 80.0, 0.0, 100.0, 0.0, 260.0, 0.0, 120.0, 0.0, 100.0, 0.0, 260.0, 0.0, 100.0, 0.0, 120.0, 0.0, 260.0, 0.0, 100.0, 0.0, 80.0, 0.0, 260.0, 80.0, 0.0, 100.0, 0.0, 260.0, 0.0, 120.0, 0.0, 100.0, 0.0, 260.0, 0.0, 100.0, 0.0, 120.0, 0.0, 260.0, 0.0, 100.0, 0.0, 80.0, 0.0, 260.0, 0.0, 0.0, 0.0, 0.0, 0.0, 0.0, 0.0, 0.0, 0.0, 0.0, 0.0, 0.0, 0.0, 0.0, 0.0, 0.0, 0.0, 0.0, 0.0, 0.0, 0.0, 0.0, 0.0, 80.0, 0.0, 100.0, 0.0, 260.0, 0.0, 120.0, 0.0, 100.0, 0.0, 260.0, 0.0, 220.0, 0.0, 240.0, 0.0, 260.0, 0.0, 100.0, 0.0, 80.0, 0.0, 260.0, 80.0, 0.0, 100.0, 0.0, 260.0, 0.0, 120.0, 0.0, 100.0, 0.0, 260.0, 0.0, 220.0, 0.0, 240.0, 0.0, 260.0, 0.0, 100.0, 0.0, 80.0, 0.0, 260.0, 80.0, 0.0, 100.0, 0.0, 260.0, 0.0, 120.0, 0.0, 100.0, 0.0, 260.0, 0.0, 220.0, 0.0, 240.0, 0.0, 260.0, 0.0, 100.0, 0.0, 80.0, 0.0, 260.0, 80.0, 0.0, 100.0, 0.0, 260.0, 0.0, 120.0, 0.0, 100.0, 0.0, 260.0, 0.0, 220.0, 0.0, 240.0, 0.0, 260.0, 0.0, 100.0, 0.0, 80.0, 0.0, 260.0, 80.0, 0.0, 100.0, 0.0, 260.0, 0.0, 120.0, 0.0, 100.0, 0.0, 260.0, 0.0, 340.0, 0.0, 360.0, 0.0, 260.0, 0.0, 100.0, 0.0, 80.0, 0.0, 260.0, 80.0, 0.0, 100.0, 0.0, 260.0, 0.0, 120.0, 0.0, 100.0, 0.0, 260.0, 0.0, 340.0, 0.0, 360.0, 0.0, 260.0, 0.0, 100.0, 0.0, 80.0, 0.0, 260.0, 80.0, 0.0, 100.0, 0.0, 260.0, 0.0, 120.0, 0.0, 100.0, 0.0, 260.0, 0.0, 340.0, 0.0, 360.0, 0.0, 260.0, 0.0, 100.0, 0.0, 80.0, 0.0, 260.0, 80.0, 0.0, 100.0, 0.0, 260.0, 0.0, 120.0, 0.0, 100.0, 0.0, 260.0, 0.0, 340.0, 0.0, 360.0, 0.0, 260.0, 0.0, 100.0, 0.0, 80.0, 0.0, 260.0, 80.0, 0.0, 100.0, 0.0, 260.0, 0.0, 240.0, 0.0, 220.0, 0.0, 260.0, 0.0, 100.0, 0.0, 120.0, 0.0, 260.0, 0.0, 100.0, 0.0, 80.0, 0.0, 260.0, 80.0, 0.0, 100.0, 0.0, 260.0, 0.0, 240.0, 0.0, 220.0, 0.0, 260.0, 0.0, 100.0, 0.0, 120.0, 0.0, 260.0, 0.0, 100.0, 0.0, 80.0, 0.0, 260.0, 80.0, 0.0, 100.0, 0.0, 260.0, 0.0, 240.0, 0.0, 220.0, 0.0, 260.0, 0.0, 100.0, 0.0, 120.0, 0.0, 260.0, 0.0, 100.0, 0.0, 80.0, 0.0, 260.0, 80.0, 0.0, 100.0, 0.0, 260.0, 0.0, 240.0, 0.0, 220.0, 0.0, 260.0, 0.0, 100.0, 0.0, 120.0, 0.0, 260.0, 0.0, 100.0, 0.0, 80.0, 0.0, 260.0, 0.0, 0.0, 0.0, 0.0, 0.0, 0.0, 0.0, 0.0, 0.0, 0.0, 0.0, 0.0, 0.0, 0.0, 0.0, 0.0, 0.0, 0.0, 0.0, 0.0, 0.0, 0.0, 0.0, 80.0, 0.0, 100.0, 0.0, 260.0, 0.0, 240.0, 0.0, 220.0, 0.0, 260.0, 0.0, 220.0, 0.0, 240.0, 0.0, 260.0, 0.0, 100.0, 0.0, 80.0, 0.0, 260.0, 80.0, 0.0, 100.0, 0.0, 260.0, 0.0, 240.0, 0.0, 220.0, 0.0, 260.0, 0.0, 220.0, 0.0, 240.0, 0.0, 260.0, 0.0, 100.0, 0.0, 80.0, 0.0, 260.0, 80.0, 0.0, 100.0, 0.0, 260.0, 0.0, 240.0, 0.0, 220.0, 0.0, 260.0, 0.0, 220.0, 0.0, 240.0, 0.0, 260.0, 0.0, 100.0, 0.0, 80.0, 0.0, 260.0, 80.0, 0.0, 100.0, 0.0, 260.0, 0.0, 240.0, 0.0, 220.0, 0.0, 260.0, 0.0, 340.0, 0.0, 360.0, 0.0, 260.0, 0.0, 100.0, 0.0, 80.0, 0.0, 260.0, 80.0, 0.0, 100.0, 0.0, 260.0, 0.0, 240.0, 0.0, 220.0, 0.0, 260.0, 0.0, 340.0, 0.0, 360.0, 0.0, 260.0, 0.0, 100.0, 0.0, 80.0, 0.0, 260.0, 80.0, 0.0, 100.0, 0.0, 260.0, 0.0, 240.0, 0.0, 220.0, 0.0, 260.0, 0.0, 340.0, 0.0, 360.0, 0.0, 260.0, 0.0, 100.0, 0.0, 80.0, 0.0, 260.0, 80.0, 0.0, 100.0, 0.0, 260.0, 0.0, 240.0, 0.0, 220.0, 0.0, 260.0, 0.0, 340.0, 0.0, 360.0, 0.0, 260.0, 0.0, 100.0, 0.0, 80.0, 0.0, 260.0, 80.0, 0.0, 100.0, 0.0, 260.0, 0.0, 240.0, 0.0, 220.0, 0.0, 260.0, 0.0, 100.0, 0.0, 120.0, 0.0, 260.0, 0.0, 100.0, 0.0, 80.0, 0.0, 260.0, 80.0, 0.0, 100.0, 0.0, 260.0, 0.0, 240.0, 0.0, 220.0, 0.0, 260.0, 0.0, 100.0, 0.0, 120.0, 0.0, 260.0, 0.0, 100.0, 0.0, 80.0, 0.0, 260.0, 80.0, 0.0, 100.0, 0.0, 260.0, 0.0, 240.0, 0.0, 220.0, 0.0, 260.0, 0.0, 100.0, 0.0, 120.0, 0.0, 260.0, 0.0, 100.0, 0.0, 80.0, 0.0, 260.0, 80.0, 0.0, 100.0, 0.0, 260.0, 0.0, 240.0, 0.0, 220.0, 0.0, 260.0, 0.0, 100.0, 0.0, 120.0, 0.0, 260.0, 0.0, 100.0, 0.0, 80.0, 0.0, 260.0, 80.0, 0.0, 100.0, 0.0, 260.0, 0.0, 240.0, 0.0, 220.0, 0.0, 260.0, 0.0, 220.0, 0.0, 240.0, 0.0, 260.0, 0.0, 100.0, 0.0, 80.0, 0.0, 260.0, 0.0, 0.0, 0.0, 0.0, 0.0, 0.0, 0.0, 0.0, 0.0, 0.0, 0.0, 0.0, 0.0, 0.0, 0.0, 0.0, 0.0, 0.0, 0.0, 0.0, 0.0, 0.0, 0.0, 80.0, 0.0, 100.0, 0.0, 260.0, 0.0, 240.0, 0.0, 220.0, 0.0, 260.0, 0.0, 220.0, 0.0, 240.0, 0.0, 260.0, 0.0, 100.0, 0.0, 80.0, 0.0, 260.0, 80.0, 0.0, 100.0, 0.0, 260.0, 0.0, 240.0, 0.0, 220.0, 0.0, 260.0, 0.0, 220.0, 0.0, 240.0, 0.0, 260.0, 0.0, 100.0, 0.0, 80.0, 0.0, 260.0, 80.0, 0.0, 100.0, 0.0, 260.0, 0.0, 240.0, 0.0, 220.0, 0.0, 260.0, 0.0, 340.0, 0.0, 360.0, 0.0, 260.0, 0.0, 100.0, 0.0, 80.0, 0.0, 260.0, 80.0, 0.0, 100.0, 0.0, 260.0, 0.0, 240.0, 0.0, 220.0, 0.0, 260.0, 0.0, 340.0, 0.0, 360.0, 0.0, 260.0, 0.0, 100.0, 0.0, 80.0, 0.0, 260.0, 80.0, 0.0, 100.0, 0.0, 260.0, 0.0, 240.0, 0.0, 220.0, 0.0, 260.0, 0.0, 340.0, 0.0, 360.0, 0.0, 260.0, 0.0, 100.0, 0.0, 80.0, 0.0, 260.0, 80.0, 0.0, 100.0, 0.0, 260.0, 0.0, 240.0, 0.0, 220.0, 0.0, 260.0, 0.0, 340.0, 0.0, 360.0, 0.0, 260.0, 0.0, 100.0, 0.0, 80.0, 0.0, 260.0, 80.0, 0.0, 100.0, 0.0, 260.0, 0.0, 240.0, 0.0, 220.0, 0.0, 260.0, 0.0, 100.0, 0.0, 120.0, 0.0, 260.0, 0.0, 100.0, 0.0, 80.0, 0.0, 260.0, 80.0, 0.0, 100.0, 0.0, 260.0, 0.0, 240.0, 0.0, 220.0, 0.0, 260.0, 0.0, 100.0, 0.0, 120.0, 0.0, 260.0, 0.0, 100.0, 0.0, 80.0, 0.0, 260.0, 80.0, 0.0, 100.0, 0.0, 260.0, 0.0, 240.0, 0.0, 220.0, 0.0, 260.0, 0.0, 100.0, 0.0, 120.0, 0.0, 260.0, 0.0, 100.0, 0.0, 80.0, 0.0, 260.0, 80.0, 0.0, 100.0, 0.0, 260.0, 0.0, 240.0, 0.0, 220.0, 0.0, 260.0, 0.0, 100.0, 0.0, 120.0, 0.0, 260.0, 0.0, 100.0, 0.0, 80.0, 0.0, 260.0, 80.0, 0.0, 100.0, 0.0, 260.0, 0.0, 240.0, 0.0, 220.0, 0.0, 260.0, 0.0, 220.0, 0.0, 240.0, 0.0, 260.0, 0.0, 100.0, 0.0, 80.0, 0.0, 260.0, 80.0, 0.0, 100.0, 0.0, 260.0, 0.0, 240.0, 0.0, 220.0, 0.0, 260.0, 0.0, 220.0, 0.0, 240.0, 0.0, 260.0, 0.0, 100.0, 0.0, 80.0, 0.0, 260.0, 0.0, 0.0, 0.0, 0.0, 0.0, 0.0, 0.0, 0.0, 0.0, 0.0, 0.0, 0.0, 0.0, 0.0, 0.0, 0.0, 0.0, 0.0, 0.0, 0.0, 0.0, 0.0, 0.0, 80.0, 0.0, 100.0, 0.0, 260.0, 0.0, 240.0, 0.0, 220.0, 0.0, 260.0, 0.0, 220.0, 0.0, 240.0, 0.0, 260.0, 0.0, 100.0, 0.0, 80.0, 0.0, 260.0, 80.0, 0.0, 100.0, 0.0, 260.0, 0.0, 240.0, 0.0, 220.0, 0.0, 260.0, 0.0, 340.0, 0.0, 360.0, 0.0, 260.0, 0.0, 100.0, 0.0, 80.0, 0.0, 260.0, 80.0, 0.0, 100.0, 0.0, 260.0, 0.0, 240.0, 0.0, 220.0, 0.0, 260.0, 0.0, 340.0, 0.0, 360.0, 0.0, 260.0, 0.0, 100.0, 0.0, 80.0, 0.0, 260.0, 80.0, 0.0, 100.0, 0.0, 260.0, 0.0, 240.0, 0.0, 220.0, 0.0, 260.0, 0.0, 340.0, 0.0, 360.0, 0.0, 260.0, 0.0, 100.0, 0.0, 80.0, 0.0, 260.0, 80.0, 0.0, 100.0, 0.0, 260.0, 0.0, 240.0, 0.0, 220.0, 0.0, 260.0, 0.0, 340.0, 0.0, 360.0, 0.0, 260.0, 0.0, 100.0, 0.0, 80.0, 0.0, 260.0, 80.0, 0.0, 100.0, 0.0, 260.0, 0.0, 240.0, 0.0, 220.0, 0.0, 260.0, 0.0, 100.0, 0.0, 120.0, 0.0, 260.0, 0.0, 100.0, 0.0, 80.0, 0.0, 260.0, 80.0, 0.0, 100.0, 0.0, 260.0, 0.0, 240.0, 0.0, 220.0, 0.0, 260.0, 0.0, 100.0, 0.0, 120.0, 0.0, 260.0, 0.0, 100.0, 0.0, 80.0, 0.0, 260.0, 80.0, 0.0, 100.0, 0.0, 260.0, 0.0, 240.0, 0.0, 220.0, 0.0, 260.0, 0.0, 100.0, 0.0, 120.0, 0.0, 260.0, 0.0, 100.0, 0.0, 80.0, 0.0, 260.0, 80.0, 0.0, 100.0, 0.0, 260.0, 0.0, 240.0, 0.0, 220.0, 0.0, 260.0, 0.0, 100.0, 0.0, 120.0, 0.0, 260.0, 0.0, 100.0, 0.0, 80.0, 0.0, 260.0, 80.0, 0.0, 100.0, 0.0, 260.0, 0.0, 240.0, 0.0, 220.0, 0.0, 260.0, 0.0, 220.0, 0.0, 240.0, 0.0, 260.0, 0.0, 100.0, 0.0, 80.0, 0.0, 260.0, 80.0, 0.0, 100.0, 0.0, 260.0, 0.0, 240.0, 0.0, 220.0, 0.0, 260.0, 0.0, 220.0, 0.0, 240.0, 0.0, 260.0, 0.0, 100.0, 0.0, 80.0, 0.0, 260.0, 80.0, 0.0, 100.0, 0.0, 260.0, 0.0, 240.0, 0.0, 220.0, 0.0, 260.0, 0.0, 220.0, 0.0, 240.0, 0.0, 260.0, 0.0, 100.0, 0.0, 80.0, 0.0, 260.0, 0.0, 0.0, 0.0, 0.0, 0.0, 0.0, 0.0, 0.0, 0.0, 0.0, 0.0, 0.0, 0.0, 0.0, 0.0, 0.0, 0.0, 0.0, 0.0, 0.0, 0.0, 0.0, 0.0, 80.0, 0.0, 100.0, 0.0, 260.0, 0.0, 240.0, 0.0, 220.0, 0.0, 260.0, 0.0, 340.0, 0.0, 360.0, 0.0, 260.0, 0.0, 100.0, 0.0, 80.0, 0.0, 260.0, 80.0, 0.0, 100.0, 0.0, 260.0, 0.0, 240.0, 0.0, 220.0, 0.0, 260.0, 0.0, 340.0, 0.0, 360.0, 0.0, 260.0, 0.0, 100.0, 0.0, 80.0, 0.0, 260.0, 80.0, 0.0, 100.0, 0.0, 260.0, 0.0, 240.0, 0.0, 220.0, 0.0, 260.0, 0.0, 340.0, 0.0, 360.0, 0.0, 260.0, 0.0, 100.0, 0.0, 80.0, 0.0, 260.0, 80.0, 0.0, 100.0, 0.0, 260.0, 0.0, 240.0, 0.0, 220.0, 0.0, 260.0, 0.0, 340.0, 0.0, 360.0, 0.0, 260.0, 0.0, 100.0, 0.0, 80.0, 0.0, 260.0, 80.0, 0.0, 100.0, 0.0, 260.0, 0.0, 360.0, 0.0, 340.0, 0.0, 260.0, 0.0, 100.0, 0.0, 120.0, 0.0, 260.0, 0.0, 100.0, 0.0, 80.0, 0.0, 260.0, 80.0, 0.0, 100.0, 0.0, 260.0, 0.0, 360.0, 0.0, 340.0, 0.0, 260.0, 0.0, 100.0, 0.0, 120.0, 0.0, 260.0, 0.0, 100.0, 0.0, 80.0, 0.0, 260.0, 80.0, 0.0, 100.0, 0.0, 260.0, 0.0, 360.0, 0.0, 340.0, 0.0, 260.0, 0.0, 100.0, 0.0, 120.0, 0.0, 260.0, 0.0, 100.0, 0.0, 80.0, 0.0, 260.0, 80.0, 0.0, 100.0, 0.0, 260.0, 0.0, 360.0, 0.0, 340.0, 0.0, 260.0, 0.0, 100.0, 0.0, 120.0, 0.0, 260.0, 0.0, 100.0, 0.0, 80.0, 0.0, 260.0, 80.0, 0.0, 100.0, 0.0, 260.0, 0.0, 360.0, 0.0, 340.0, 0.0, 260.0, 0.0, 220.0, 0.0, 240.0, 0.0, 260.0, 0.0, 100.0, 0.0, 80.0, 0.0, 260.0, 80.0, 0.0, 100.0, 0.0, 260.0, 0.0, 360.0, 0.0, 340.0, 0.0, 260.0, 0.0, 220.0, 0.0, 240.0, 0.0, 260.0, 0.0, 100.0, 0.0, 80.0, 0.0, 260.0, 80.0, 0.0, 100.0, 0.0, 260.0, 0.0, 360.0, 0.0, 340.0, 0.0, 260.0, 0.0, 220.0, 0.0, 240.0, 0.0, 260.0, 0.0, 100.0, 0.0, 80.0, 0.0, 260.0, 80.0, 0.0, 100.0, 0.0, 260.0, 0.0, 360.0, 0.0, 340.0, 0.0, 260.0, 0.0, 220.0, 0.0, 240.0, 0.0, 260.0, 0.0, 100.0, 0.0, 80.0, 0.0, 260.0, 0.0, 0.0, 0.0, 0.0, 0.0, 0.0, 0.0, 0.0, 0.0, 0.0, 0.0, 0.0, 0.0, 0.0, 0.0, 0.0, 0.0, 0.0, 0.0, 0.0, 0.0, 0.0, 0.0, 80.0, 0.0, 100.0, 0.0, 260.0, 0.0, 360.0, 0.0, 340.0, 0.0, 260.0, 0.0, 340.0, 0.0, 360.0, 0.0, 260.0, 0.0, 100.0, 0.0, 80.0, 0.0, 260.0, 80.0, 0.0, 100.0, 0.0, 260.0, 0.0, 360.0, 0.0, 340.0, 0.0, 260.0, 0.0, 340.0, 0.0, 360.0, 0.0, 260.0, 0.0, 100.0, 0.0, 80.0, 0.0, 260.0, 80.0, 0.0, 100.0, 0.0, 260.0, 0.0, 360.0, 0.0, 340.0, 0.0, 260.0, 0.0, 340.0, 0.0, 360.0, 0.0, 260.0, 0.0, 100.0, 0.0, 80.0, 0.0, 260.0, 80.0, 0.0, 100.0, 0.0, 260.0, 0.0, 360.0, 0.0, 340.0, 0.0, 260.0, 0.0, 100.0, 0.0, 120.0, 0.0, 260.0, 0.0, 100.0, 0.0, 80.0, 0.0, 260.0, 80.0, 0.0, 100.0, 0.0, 260.0, 0.0, 360.0, 0.0, 340.0, 0.0, 260.0, 0.0, 100.0, 0.0, 120.0, 0.0, 260.0, 0.0, 100.0, 0.0, 80.0, 0.0, 260.0, 80.0, 0.0, 100.0, 0.0, 260.0, 0.0, 360.0, 0.0, 340.0, 0.0, 260.0, 0.0, 100.0, 0.0, 120.0, 0.0, 260.0, 0.0, 100.0, 0.0, 80.0, 0.0, 260.0, 80.0, 0.0, 100.0, 0.0, 260.0, 0.0, 360.0, 0.0, 340.0, 0.0, 260.0, 0.0, 100.0, 0.0, 120.0, 0.0, 260.0, 0.0, 100.0, 0.0, 80.0, 0.0, 260.0, 80.0, 0.0, 100.0, 0.0, 260.0, 0.0, 360.0, 0.0, 340.0, 0.0, 260.0, 0.0, 220.0, 0.0, 240.0, 0.0, 260.0, 0.0, 100.0, 0.0, 80.0, 0.0, 260.0, 80.0, 0.0, 100.0, 0.0, 260.0, 0.0, 360.0, 0.0, 340.0, 0.0, 260.0, 0.0, 220.0, 0.0, 240.0, 0.0, 260.0, 0.0, 100.0, 0.0, 80.0, 0.0, 260.0, 80.0, 0.0, 100.0, 0.0, 260.0, 0.0, 360.0, 0.0, 340.0, 0.0, 260.0, 0.0, 220.0, 0.0, 240.0, 0.0, 260.0, 0.0, 100.0, 0.0, 80.0, 0.0, 260.0, 80.0, 0.0, 100.0, 0.0, 260.0, 0.0, 360.0, 0.0, 340.0, 0.0, 260.0, 0.0, 220.0, 0.0, 240.0, 0.0, 260.0, 0.0, 100.0, 0.0, 80.0, 0.0, 260.0, 80.0, 0.0, 100.0, 0.0, 260.0, 0.0, 360.0, 0.0, 340.0, 0.0, 260.0, 0.0, 340.0, 0.0, 360.0, 0.0, 260.0, 0.0, 100.0, 0.0, 80.0, 0.0, 260.0, 0.0, 0.0, 0.0, 0.0, 0.0, 0.0, 0.0, 0.0, 0.0, 0.0, 0.0, 0.0, 0.0, 0.0, 0.0, 0.0, 0.0, 0.0, 0.0, 0.0, 0.0, 0.0, 0.0, 80.0, 0.0, 100.0, 0.0, 260.0, 0.0, 360.0, 0.0, 340.0, 0.0, 260.0, 0.0, 340.0, 0.0, 360.0, 0.0, 260.0, 0.0, 100.0, 0.0, 80.0, 0.0, 260.0, 80.0, 0.0, 100.0, 0.0, 260.0, 0.0, 360.0, 0.0, 340.0, 0.0, 260.0, 0.0, 340.0, 0.0, 360.0, 0.0, 260.0, 0.0, 100.0, 0.0, 80.0, 0.0, 260.0, 80.0, 0.0, 100.0, 0.0, 260.0, 0.0, 360.0, 0.0, 340.0, 0.0, 260.0, 0.0, 100.0, 0.0, 120.0, 0.0, 260.0, 0.0, 100.0, 0.0, 80.0, 0.0, 260.0, 80.0, 0.0, 100.0, 0.0, 260.0, 0.0, 360.0, 0.0, 340.0, 0.0, 260.0, 0.0, 100.0, 0.0, 120.0, 0.0, 260.0, 0.0, 100.0, 0.0, 80.0, 0.0, 260.0, 80.0, 0.0, 100.0, 0.0, 260.0, 0.0, 360.0, 0.0, 340.0, 0.0, 260.0, 0.0, 100.0, 0.0, 120.0, 0.0, 260.0, 0.0, 100.0, 0.0, 80.0, 0.0, 260.0, 80.0, 0.0, 100.0, 0.0, 260.0, 0.0, 360.0, 0.0, 340.0, 0.0, 260.0, 0.0, 100.0, 0.0, 120.0, 0.0, 260.0, 0.0, 100.0, 0.0, 80.0, 0.0, 260.0, 80.0, 0.0, 100.0, 0.0, 260.0, 0.0, 360.0, 0.0, 340.0, 0.0, 260.0, 0.0, 220.0, 0.0, 240.0, 0.0, 260.0, 0.0, 100.0, 0.0, 80.0, 0.0, 260.0, 80.0, 0.0, 100.0, 0.0, 260.0, 0.0, 360.0, 0.0, 340.0, 0.0, 260.0, 0.0, 220.0, 0.0, 240.0, 0.0, 260.0, 0.0, 100.0, 0.0, 80.0, 0.0, 260.0, 80.0, 0.0, 100.0, 0.0, 260.0, 0.0, 360.0, 0.0, 340.0, 0.0, 260.0, 0.0, 220.0, 0.0, 240.0, 0.0, 260.0, 0.0, 100.0, 0.0, 80.0, 0.0, 260.0, 80.0, 0.0, 100.0, 0.0, 260.0, 0.0, 360.0, 0.0, 340.0, 0.0, 260.0, 0.0, 220.0, 0.0, 240.0, 0.0, 260.0, 0.0, 100.0, 0.0, 80.0, 0.0, 260.0, 80.0, 0.0, 100.0, 0.0, 260.0, 0.0, 360.0, 0.0, 340.0, 0.0, 260.0, 0.0, 340.0, 0.0, 360.0, 0.0, 260.0, 0.0, 100.0, 0.0, 80.0, 0.0, 260.0, 80.0, 0.0, 100.0, 0.0, 260.0, 0.0, 360.0, 0.0, 340.0, 0.0, 260.0, 0.0, 340.0, 0.0, 360.0, 0.0, 260.0, 0.0, 100.0, 0.0, 80.0, 0.0, 260.0, 0.0, 0.0, 0.0, 0.0, 0.0, 0.0, 0.0, 0.0, 0.0, 0.0, 0.0, 0.0, 0.0, 0.0, 0.0, 0.0, 0.0, 0.0, 0.0, 0.0, 0.0, 0.0, 0.0, 80.0, 0.0, 100.0, 0.0, 260.0, 0.0, 360.0, 0.0, 340.0, 0.0, 260.0, 0.0, 340.0, 0.0, 360.0, 0.0, 260.0, 0.0, 100.0, 0.0, 80.0, 0.0, 260.0, 80.0, 0.0, 100.0, 0.0, 260.0, 0.0, 360.0, 0.0, 340.0, 0.0, 260.0, 0.0, 100.0, 0.0, 120.0, 0.0, 260.0, 0.0, 100.0, 0.0, 80.0, 0.0, 260.0, 80.0, 0.0, 100.0, 0.0, 260.0, 0.0, 360.0, 0.0, 340.0, 0.0, 260.0, 0.0, 100.0, 0.0, 120.0, 0.0, 260.0, 0.0, 100.0, 0.0, 80.0, 0.0, 260.0, 80.0, 0.0, 100.0, 0.0, 260.0, 0.0, 360.0, 0.0, 340.0, 0.0, 260.0, 0.0, 100.0, 0.0, 120.0, 0.0, 260.0, 0.0, 100.0, 0.0, 80.0, 0.0, 260.0, 80.0, 0.0, 100.0, 0.0, 260.0, 0.0, 360.0, 0.0, 340.0, 0.0, 260.0, 0.0, 100.0, 0.0, 120.0, 0.0, 260.0, 0.0, 100.0, 0.0, 80.0, 0.0, 260.0, 80.0, 0.0, 100.0, 0.0, 260.0, 0.0, 360.0, 0.0, 340.0, 0.0, 260.0, 0.0, 220.0, 0.0, 240.0, 0.0, 260.0, 0.0, 100.0, 0.0, 80.0, 0.0, 260.0, 80.0, 0.0, 100.0, 0.0, 260.0, 0.0, 360.0, 0.0, 340.0, 0.0, 260.0, 0.0, 220.0, 0.0, 240.0, 0.0, 260.0, 0.0, 100.0, 0.0, 80.0, 0.0, 260.0, 80.0, 0.0, 100.0, 0.0, 260.0, 0.0, 360.0, 0.0, 340.0, 0.0, 260.0, 0.0, 220.0, 0.0, 240.0, 0.0, 260.0, 0.0, 100.0, 0.0, 80.0, 0.0, 260.0, 80.0, 0.0, 100.0, 0.0, 260.0, 0.0, 360.0, 0.0, 340.0, 0.0, 260.0, 0.0, 220.0, 0.0, 240.0, 0.0, 260.0, 0.0, 100.0, 0.0, 80.0, 0.0, 260.0, 80.0, 0.0, 100.0, 0.0, 260.0, 0.0, 360.0, 0.0, 340.0, 0.0, 260.0, 0.0, 340.0, 0.0, 360.0, 0.0, 260.0, 0.0, 100.0, 0.0, 80.0, 0.0, 260.0, 80.0, 0.0, 100.0, 0.0, 260.0, 0.0, 360.0, 0.0, 340.0, 0.0, 260.0, 0.0, 340.0, 0.0, 360.0, 0.0, 260.0, 0.0, 100.0, 0.0, 80.0, 0.0, 260.0, 80.0, 0.0, 100.0, 0.0, 260.0, 0.0, 360.0, 0.0, 340.0, 0.0, 260.0, 0.0, 340.0, 0.0, 360.0, 0.0, 260.0, 0.0, 100.0, 0.0, 80.0, 0.0, 260.0];
    TG_STORE_TRAVEL : ARRAY[1..12, 1..12] OF REAL := [0.0, 0.0, 0.0, 0.0, 0.0, 120.0, 0.0, 0.0, 0.0, 0.0, 0.0, 665.0, 0.0, 0.0, 0.0, 0.0, 0.0, 240.0, 0.0, 0.0, 0.0, 0.0, 0.0, 665.0, 0.0, 0.0, 0.0, 0.0, 0.0, 360.0, 0.0, 0.0, 0.0, 0.0, 0.0, 665.0, 0.0, 0.0, 0.0, 0.0, 0.0, 480.0, 0.0, 0.0, 0.0, 0.0, 0.0, 665.0, 0.0, 0.0, 0.0, 0.0, 0.0, 120.0, 0.0, 0.0, 0.0, 0.0, 0.0, 665.0, 0.0, 0.0, 0.0, 0.0, 0.0, 240.0, 0.0, 0.0, 0.0, 0.0, 0.0, 665.0, 0.0, 0.0, 0.0, 0.0, 0.0, 360.0, 0.0, 0.0, 0.0, 0.0, 0.0, 665.0, 0.0, 0.0, 0.0, 0.0, 0.0, 480.0, 0.0, 0.0, 0.0, 0.0, 0.0, 665.0, 0.0, 0.0, 0.0, 0.0, 0.0, 120.0, 0.0, 0.0, 0.0, 0.0, 0.0, 665.0, 0.0, 0.0, 0.0, 0.0, 0.0, 240.0, 0.0, 0.0, 0.0, 0.0, 0.0, 665.0, 0.0, 0.0, 0.0, 0.0, 0.0, 360.0, 0.0, 0.0, 0.0, 0.0, 0.0, 665.0, 0.0, 0.0, 0.0, 0.0, 0.0, 480.0, 0.0, 0.0, 0.0, 0.0, 0.0, 665.0];
    TG_STORE_LIFT : ARRAY[1..12, 1..12] OF REAL := [80.0, 0.0, 100.0, 0.0, 260.0, 0.0, 120.0, 0.0, 100.0, 0.0, 260.0, 0.0, 80.0, 0.0, 100.0, 0.0, 260.0, 0.0, 120.0, 0.0, 100.0, 0.0, 260.0, 0.0, 80.0, 0.0, 100.0, 0.0, 260.0, 0.0, 120.0, 0.0, 100.0, 0.0, 260.0, 0.0, 80.0, 0.0, 100.0, 0.0, 260.0, 0.0, 120.0, 0.0, 100.0, 0.0, 260.0, 0.0, 80.0, 0.0, 100.0, 0.0, 260.0, 0.0, 240.0, 0.0, 220.0, 0.0, 260.0, 0.0, 80.0, 0.0, 100.0, 0.0, 260.0, 0.0, 240.0, 0.0, 220.0, 0.0, 260.0, 0.0, 80.0, 0.0, 100.0, 0.0, 260.0, 0.0, 240.0, 0.0, 220.0, 0.0, 260.0, 0.0, 80.0, 0.0, 100.0, 0.0, 260.0, 0.0, 240.0, 0.0, 220.0, 0.0, 260.0, 0.0, 80.0, 0.0, 100.0, 0.0, 260.0, 0.0, 360.0, 0.0, 340.0, 0.0, 260.0, 0.0, 80.0, 0.0, 100.0, 0.0, 260.0, 0.0, 360.0, 0.0, 340.0, 0.0, 260.0, 0.0, 80.0, 0.0, 100.0, 0.0, 260.0, 0.0, 360.0, 0.0, 340.0, 0.0, 260.0, 0.0, 80.0, 0.0, 100.0, 0.0, 260.0, 0.0, 360.0, 0.0, 340.0, 0.0, 260.0, 0.0];
    TG_FETCH_EMPTY_TRAVEL : ARRAY[1..12, 1..12] OF REAL := [120.0, 0.0, 0.0, 0.0, 0.0, 0.0, 665.0, 0.0, 0.0, 0.0, 0.0, 0.0, 240.0, 0.0, 0.0, 0.0, 0.0, 0.0, 665.0, 0.0, 0.0, 0.0, 0.0, 0.0, 360.0, 0.0, 0.0, 0.0, 0.0, 0.0, 665.0, 0.0, 0.0, 0.0, 0.0, 0.0, 480.0, 0.0, 0.0, 0.0, 0.0, 0.0, 665.0, 0.0, 0.0, 0.0, 0.0, 0.0, 120.0, 0.0, 0.0, 0.0, 0.0, 0.0, 665.0, 0.0, 0.0, 0.0, 0.0, 0.0, 240.0, 0.0, 0.0, 0.0, 0.0, 0.0, 665.0, 0.0, 0.0, 0.0, 0.0, 0.0, 360.0, 0.0, 0.0, 0.0, 0.0, 0.0, 665.0, 0.0, 0.0, 0.0, 0.0, 0.0, 480.0, 0.0, 0.0, 0.0, 0.0, 0.0, 665.0, 0.0, 0.0, 0.0, 0.0, 0.0, 120.0, 0.0, 0.0, 0.0, 0.0, 0.0, 665.0, 0.0, 0.0, 0.0, 0.0, 0.0, 240.0, 0.0, 0.0, 0.0, 0.0, 0.0, 665.0, 0.0, 0.0, 0.0, 0.0, 0.0, 360.0, 0.0, 0.0, 0.0, 0.0, 0.0, 665.0, 0.0, 0.0, 0.0, 0.0, 0.0, 480.0, 0.0, 0.0, 0.0, 0.0, 0.0, 665.0, 0.0, 0.0, 0.0, 0.0, 0.0];
    TG_FETCH_EMPTY_LIFT : ARRAY[1..12, 1..12] OF REAL := [0.0, 100.0, 0.0, 120.0, 0.0, 260.0, 0.0, 100.0, 0.0, 80.0, 0.0, 260.0, 0.0, 100.0, 0.0, 120.0, 0.0, 260.0, 0.0, 100.0, 0.0, 80.0, 0.0, 260.0, 0.0, 100.0, 0.0, 120.0, 0.0, 260.0, 0.0, 100.0, 0.0, 80.0, 0.0, 260.0, 0.0, 100.0, 0.0, 120.0, 0.0, 260.0, 0.0, 100.0, 0.0, 80.0, 0.0, 260.0, 0.0, 220.0, 0.0, 240.0, 0.0, 260.0, 0.0, 100.0, 0.0, 80.0, 0.0, 260.0, 0.0, 220.0, 0.0, 240.0, 0.0, 260.0, 0.0, 100.0, 0.0, 80.0, 0.0, 260.0, 0.0, 220.0, 0.0, 240.0, 0.0, 260.0, 0.0, 100.0, 0.0, 80.0, 0.0, 260.0, 0.0, 220.0, 0.0, 240.0, 0.0, 260.0, 0.0, 100.0, 0.0, 80.0, 0.0, 260.0, 0.0, 340.0, 0.0, 360.0, 0.0, 260.0, 0.0, 100.0, 0.0, 80.0, 0.0, 260.0, 0.0, 340.0, 0.0, 360.0, 0.0, 260.0, 0.0, 100.0, 0.0, 80.0, 0.0, 260.0, 0.0, 340.0, 0.0, 360.0, 0.0, 260.0, 0.0, 100.0, 0.0, 80.0, 0.0, 260.0, 0.0, 340.0, 0.0, 360.0, 0.0, 260.0, 0.0, 100.0, 0.0, 80.0, 0.0, 260.0];
    TG_RETRIEVE_TRAVEL : ARRAY[1..12, 1..12] OF REAL := [120.0, 0.0, 0.0, 0.0, 0.0, 0.0, 665.0, 0.0, 0.0, 0.0, 0.0, 0.0, 240.0, 0.0, 0.0, 0.0, 0.0, 0.0, 665.0, 0.0, 0.0, 0.0, 0.0, 0.0, 360.0, 0.0, 0.0, 0.0, 0.0, 0.0, 665.0, 0.0, 0.0, 0.0, 0.0, 0.0, 480.0, 0.0, 0.0, 0.0, 0.0, 0.0, 665.0, 0.0, 0.0, 0.0, 0.0, 0.0, 120.0, 0.0, 0.0, 0.0, 0.0, 0.0, 665.0, 0.0, 0.0, 0.0, 0.0, 0.0, 240.0, 0.0, 0.0, 0.0, 0.0, 0.0, 665.0, 0.0, 0.0, 0.0, 0.0, 0.0, 360.0, 0.0, 0.0, 0.0, 0.0, 0.0, 665.0, 0.0, 0.0, 0.0, 0.0, 0.0, 480.0, 0.0, 0.0, 0.0, 0.0, 0.0, 665.0, 0.0, 0.0, 0.0, 0.0, 0.0, 120.0, 0.0, 0.0, 0.0, 0.0, 0.0, 665.0, 0.0, 0.0, 0.0, 0.0, 0.0, 240.0, 0.0, 0.0, 0.0, 0.0, 0.0, 665.0, 0.0, 0.0, 0.0, 0.0, 0.0, 360.0, 0.0, 0.0, 0.0, 0.0, 0.0, 665.0, 0.0, 0.0, 0.0, 0.0, 0.0, 480.0, 0.0, 0.0, 0.0, 0.0, 0.0, 665.0, 0.0, 0.0, 0.0, 0.0, 0.0];
    TG_RETRIEVE_LIFT : ARRAY[1..12, 1..12] OF REAL := [0.0, 100.0, 0.0, 120.0, 0.0, 260.0, 0.0, 100.0, 0.0, 80.0, 0.0, 260.0, 0.0, 100.0, 0.0, 120.0, 0.0, 260.0, 0.0, 100.0, 0.0, 80.0, 0.0, 260.0, 0.0, 100.0, 0.0, 120.0, 0.0, 260.0, 0.0, 100.0, 0.0, 80.0, 0.0, 260.0, 0.0, 100.0, 0.0, 120.0, 0.0, 260.0, 0.0, 100.0, 0.0, 80.0, 0.0, 260.0, 0.0, 220.0, 0.0, 240.0, 0.0, 260.0, 0.0, 100.0, 0.0, 80.0, 0.0, 260.0, 0.0, 220.0, 0.0, 240.0, 0.0, 260.0, 0.0, 100.0, 0.0, 80.0, 0.0, 260.0, 0.0, 220.0, 0.0, 240.0, 0.0, 260.0, 0.0, 100.0, 0.0, 80.0, 0.0, 260.0, 0.0, 220.0, 0.0, 240.0, 0.0, 260.0, 0.0, 100.0, 0.0, 80.0, 0.0, 260.0, 0.0, 340.0, 0.0, 360.0, 0.0, 260.0, 0.0, 100.0, 0.0, 80.0, 0.0, 260.0, 0.0, 340.0, 0.0, 360.0, 0.0, 260.0, 0.0, 100.0, 0.0, 80.0, 0.0, 260.0, 0.0, 340.0, 0.0, 360.0, 0.0, 260.0, 0.0, 100.0, 0.0, 80.0, 0.0, 260.0, 0.0, 340.0, 0.0, 360.0, 0.0, 260.0, 0.0, 100.0, 0.0, 80.0, 0.0, 260.0];
    WD_STORE_RETRIEVE : ARRAY[1..143, 1..23] OF TIME := [T#2300MS, T#1700MS, T#1100MS, T#1700MS, T#2100MS, T#6000MS, T#1900MS, T#1700MS, T#1100MS, T#1700MS, T#2100MS, T#4100MS, T#2100MS, T#1700MS, T#1100MS, T#1700MS, T#1900MS, T#6000MS, T#2100MS, T#1700MS, T#1100MS, T#1700MS, T#2300MS, T#2300MS, T#1700MS, T#1100MS, T#1700MS, T#2100MS, T#6000MS, T#1900MS, T#1700MS, T#1100MS, T#1700MS, T#2100MS, T#1700MS, T#2100MS, T#1700MS, T#1100MS, T#1700MS, T#1900MS, T#4800MS, T#2100MS, T#1700MS, T#1100MS, T#1700MS, T#2300MS, T#2300MS, T#1700MS, T#1100MS, T#1700MS, T#2100MS, T#6000MS, T#1900MS, T#1700MS, T#1100MS, T#1700MS, T#2100MS, T#2900MS, T#2100MS, T#1700MS, T#1100MS, T#1700MS, T#1900MS, T#3500MS, T#2100MS, T#1700MS, T#1100MS, T#1700MS, T#2300MS, T#2300MS, T#1700MS, T#1100MS, T#1700MS, T#2100MS, T#6000MS, T#1900MS, T#1700MS, T#1100MS, T#1700MS, T#2100MS, T#4100MS, T#2100MS, T#1700MS, T#1100MS, T#1700MS, T#1900MS, T#2400MS, T#2100MS, T#1700MS, T#1100MS, T#1700MS, T#2300MS, T#2300MS, T#1700MS, T#1100MS, T#1700MS, T#2100MS, T#6000MS, T#1900MS, T#1700MS, T#1100MS, T#1700MS, T#2100MS, T#600MS, T#1100MS, T#1700MS, T#1100MS, T#1700MS, T#1100MS, T#6000MS, T#2100MS, T#1700MS, T#1100MS, T#1700MS, T#2300MS, T#2300MS, T#1700MS, T#1100MS, T#1700MS, T#2100MS, T#6000MS, T#1900MS, T#1700MS, T#1100MS, T#1700MS, T#2100MS, T#1700MS, T#1100MS, T#1700MS, T#1100MS, T#1700MS, T#1100MS, T#4800MS, T#2100MS, T#1700MS, T#1100MS, T#1700MS, T#2300MS, T#2300MS, T#1700MS, T#1100MS, T#1700MS, T#2100MS, T#6000MS, T#1900MS, T#1700MS, T#1100MS, T#1700MS, T#2100MS, T#2900MS, T#1100MS, T#1700MS, T#1100MS, T#1700MS, T#1100MS, T#3500MS, T#2100MS, T#1700MS, T#1100MS, T#1700MS, T#2300MS, T#2300MS, T#1700MS, T#1100MS, T#1700MS, T#2100MS, T#6000MS, T#1900MS, T#1700MS, T#1100MS, T#1700MS, T#2100MS, T#4100MS, T#1100MS, T#1700MS, T#1100MS, T#1700MS, T#1100MS, T#2400MS, T#2100MS, T#1700MS, T#1100MS, T#1700MS, T#2300MS, T#2300MS, T#1700MS, T#1100MS, T#1700MS, T#2100MS, T#6000MS, T#1900MS, T#1700MS, T#1100MS, T#1700MS, T#2100MS, T#600MS, T#1300MS, T#1700MS, T#1100MS, T#1700MS, T#1500MS, T#6000MS, T#2100MS, T#1700MS, T#1100MS, T#1700MS, T#2300MS, T#2300MS, T#1700MS, T#1100MS, T#1700MS, T#2100MS, T#6000MS, T#1900MS, T#1700MS, T#1100MS, T#1700MS, T#2100MS, T#1700MS, T#1300MS, T#1700MS, T#1100MS, T#1700MS, T#1500MS, T#4800MS, T#2100MS, T#1700MS, T#1100MS, T#1700MS, T#2300MS, T#2300MS, T#1700MS, T#1100MS, T#1700MS, T#2100MS, T#6000MS, T#1900MS, T#1700MS, T#1100MS, T#1700MS, T#2100MS, T#2900MS, T#1300MS, T#1700MS, T#1100MS, T#1700MS, T#1500MS, T#3500MS, T#2100MS, T#1700MS, T#1100MS, T#1700MS, T#2300MS, T#2300MS, T#1700MS, T#1100MS, T#1700MS, T#2100MS, T#6000MS, T#1900MS, T#1700MS, T#1100MS, T#1700MS, T#2100MS, T#4100MS, T#1300MS, T#1700MS, T#1100MS, T#1700MS, T#1500MS, T#2400MS, T#2100MS, T#1700MS, T#1100MS, T#1700MS, T#2300MS, T#2300MS, T#1700MS, T#1100MS, T#1700MS, T#2100MS, T#4800MS, T#1900MS, T#1700MS, T#1100MS, T#1700MS, T#2100MS, T#1700MS, T#2100MS, T#1700MS, T#1100MS, T#1700MS, T#1900MS, T#6000MS, T#2100MS, T#1700MS, T#1100MS, T#1700MS, T#2300MS, T#2300MS, T#1700MS, T#1100MS, T#1700MS, T#2100MS, T#6000MS, T#1900MS, T#1700MS, T#1100MS, T#1700MS, T#2100MS, T#4100MS, T#2100MS, T#1700MS, T#1100MS, T#1700MS, T#1900MS, T#6000MS, T#2100MS, T#1700MS, T#1100MS, T#1700MS, T#2300MS, T#2300MS, T#1700MS, T#1100MS, T#1700MS, T#2100MS, T#4800MS, T#1900MS, T#1700MS, T#1100MS, T#1700MS, T#2100MS, T#1700MS, T#2100MS, T#1700MS, T#1100MS, T#1700MS, T#1900MS, T#3500MS, T#2100MS, T#1700MS, T#1100MS, T#1700MS, T#2300MS, T#2300MS, T#1700MS, T#1100MS, T#1700MS, T#2100MS, T#4800MS, T#1900MS, T#1700MS, T#1100MS, T#1700MS, T#2100MS, T#2900MS, T#2100MS, T#1700MS, T#1100MS, T#1700MS, T#1900MS, T#2400MS, T#2100MS, T#1700MS, T#1100MS, T#1700MS, T#2300MS, T#2300MS, T#1700MS, T#1100MS, T#1700MS, T#2100MS, T#4800MS, T#1900MS, T#1700MS, T#1100MS, T#1700MS, T#2100MS, T#1700MS, T#1100MS, T#1700MS, T#1100MS, T#1700MS, T#1100MS, T#6000MS, T#2100MS, T#1700MS, T#1100MS, T#1700MS, T#2300MS, T#2300MS, T#1700MS, T#1100MS, T#1700MS, T#2100MS, T#4800MS, T#1900MS, T#1700MS, T#1100MS, T#1700MS, T#2100MS, T#600MS, T#1100MS, T#1700MS, T#1100MS, T#1700MS, T#1100MS, T#4800MS, T#2100MS, T#1700MS, T#1100MS, T#1700MS, T#2300MS, T#2300MS, T#1700MS, T#1100MS, T#1700MS, T#2100MS, T#4800MS, T#1900MS, T#1700MS, T#1100MS, T#1700MS, T#2100MS, T#1700MS, T#1100MS, T#1700MS, T#1100MS, T#1700MS, T#1100MS, T#3500MS, T#2100MS, T#1700MS, T#1100MS, T#1700MS, T#2300MS, T#2300MS, T#1700MS, T#1100MS, T#1700MS, T#2100MS, T#4800MS, T#1900MS, T#1700MS, T#1100MS, T#1700MS, T#2100MS, T#2900MS, T#1100MS, T#1700MS, T#1100MS, T#1700MS, T#1100MS, T#2400MS, T#2100MS, T#1700MS, T#1100MS, T#1700MS, T#2300MS, T#2300MS, T#1700MS, T#1100MS, T#1700MS, T#2100MS, T#4800MS, T#1900MS, T#1700MS, T#1100MS, T#1700MS, T#2100MS, T#1700MS, T#1300MS, T#1700MS, T#1100MS, T#1700MS, T#1500MS, T#6000MS, T#2100MS, T#1700MS, T#1100MS, T#1700MS, T#2300MS, T#2300MS, T#1700MS, T#1100MS, T#1700MS, T#2100MS, T#4800MS, T#1900MS, T#1700MS, T#1100MS, T#1700MS, T#2100MS, T#600MS, T#1300MS, T#1700MS, T#1100MS, T#1700MS, T#1500MS, T#4800MS, T#2100MS, T#1700MS, T#1100MS, T#1700MS, T#2300MS, T#2300MS, T#1700MS, T#1100MS, T#1700MS, T#2100MS, T#4800MS, T#1900MS, T#1700MS, T#1100MS, T#1700MS, T#2100MS, T#1700MS, T#1300MS, T#1700MS, T#1100MS, T#1700MS, T#1500MS, T#3500MS, T#2100MS, T#1700MS, T#1100MS, T#1700MS, T#2300MS, T#2300MS, T#1700MS, T#1100MS, T#1700MS, T#2100MS, T#4800MS, T#1900MS, T#1700MS, T#1100MS, T#1700MS, T#2100MS, T#2900MS, T#1300MS, T#1700MS, T#1100MS, T#1700MS, T#1500MS, T#2400MS, T#2100MS, T#1700MS, T#1100MS, T#1700MS, T#2300MS, T#2300MS, T#1700MS, T#1100MS, T#1700MS, T#2100MS, T#3500MS, T#1900MS, T#1700MS, T#1100MS, T#1700MS, T#2100MS, T#2900MS, T#2100MS, T#1700MS, T#1100MS, T#1700MS, T#1900MS, T#6000MS, T#2100MS, T#1700MS, T#1100MS, T#1700MS, T#2300MS, T#2300MS, T#1700MS, T#1100MS, T#1700MS, T#2100MS, T#3500MS, T#1900MS, T#1700MS, T#1100MS, T#1700MS, T#2100MS, T#1700MS, T#2100MS, T#1700MS, T#1100MS, T#1700MS, T#1900MS, T#4800MS, T#2100MS, T#1700MS, T#1100MS, T#1700MS, T#2300MS, T#2300MS, T#1700MS, T#1100MS, T#1700MS, T#2100MS, T#6000MS, T#1900MS, T#1700MS, T#1100MS, T#1700MS, T#2100MS, T#4100MS, T#2100MS, T#1700MS, T#1100MS, T#1700MS, T#1900MS, T#6000MS, T#2100MS, T#1700MS, T#1100MS, T#1700MS, T#2300MS, T#2300MS, T#1700MS, T#1100MS, T#1700MS, T#2100MS, T#3500MS, T#1900MS, T#1700MS, T#1100MS, T#1700MS, T#2100MS, T#1700MS, T#2100MS, T#1700MS, T#1100MS, T#1700MS, T#1900MS, T#2400MS, T#2100MS, T#1700MS, T#1100MS, T#1700MS, T#2300MS, T#2300MS, T#1700MS, T#1100MS, T#1700MS, T#2100MS, T#3500MS, T#1900MS, T#1700MS, T#1100MS, T#1700MS, T#2100MS, T#2900MS, T#1100MS, T#1700MS, T#1100MS, T#1700MS, T#1100MS, T#6000MS, T#2100MS, T#1700MS, T#1100MS, T#1700MS, T#2300MS, T#2300MS, T#1700MS, T#1100MS, T#1700MS, T#2100MS, T#3500MS, T#1900MS, T#1700MS, T#1100MS, T#1700MS, T#2100MS, T#1700MS, T#1100MS, T#1700MS, T#1100MS, T#1700MS, T#1100MS, T#4800MS, T#2100MS, T#1700MS, T#1100MS, T#1700MS, T#2300MS, T#2300MS, T#1700MS, T#1100MS, T#1700MS, T#2100MS, T#3500MS, T#1900MS, T#1700MS, T#1100MS, T#1700MS, T#2100MS, T#600MS, T#1100MS, T#1700MS, T#1100MS, T#1700MS, T#1100MS, T#3500MS, T#2100MS, T#1700MS, T#1100MS, T#1700MS, T#2300MS, T#2300MS, T#1700MS, T#1100MS, T#1700MS, T#2100MS, T#3500MS, T#1900MS, T#1700MS, T#1100MS, T#1700MS, T#2100MS, T#1700MS, T#1100MS, T#1700MS, T#1100MS, T#1700MS, T#1100MS, T#2400MS, T#2100MS, T#1700MS, T#1100MS, T#1700MS, T#2300MS, T#2300MS, T#1700MS, T#1100MS, T#1700MS, T#2100MS, T#3500MS, T#1900MS, T#1700MS, T#1100MS, T#1700MS, T#2100MS, T#2900MS, T#1300MS, T#1700MS, T#1100MS, T#1700MS, T#1500MS, T#6000MS, T#2100MS, T#1700MS, T#1100MS, T#1700MS, T#2300MS, T#2300MS, T#1700MS, T#1100MS, T#1700MS, T#2100MS, T#3500MS, T#1900MS, T#1700MS, T#1100MS, T#1700MS, T#2100MS, T#1700MS, T#1300MS, T#1700MS, T#1100MS, T#1700MS, T#1500MS, T#4800MS, T#2100MS, T#1700MS, T#1100MS, T#1700MS, T#2300MS, T#2300MS, T#1700MS, T#1100MS, T#1700MS, T#2100MS, T#3500MS, T#1900MS, T#1700MS, T#1100MS, T#1700MS, T#2100MS, T#600MS, T#1300MS, T#1700MS, T#1100MS, T#1700MS, T#1500MS, T#3500MS, T#2100MS, T#1700MS, T#1100MS, T#1700MS, T#2300MS, T#2300MS, T#1700MS, T#1100MS, T#1700MS, T#2100MS, T#3500MS, T#1900MS, T#1700MS, T#1100MS, T#1700MS, T#2100MS, T#1700MS, T#1300MS, T#1700MS, T#1100MS, T#1700MS, T#1500MS, T#2400MS, T#2100MS, T#1700MS, T#1100MS, T#1700MS, T#2300MS, T#2300MS, T#1700MS, T#1100MS, T#1700MS, T#2100MS, T#2400MS, T#1900MS, T#1700MS, T#1100MS, T#1700MS, T#2100MS, T#4100MS, T#2100MS, T#1700MS, T#1100MS, T#1700MS, T#1900MS, T#6000MS, T#2100MS, T#1700MS, T#1100MS, T#1700MS, T#2300MS, T#2300MS, T#1700MS, T#1100MS, T#1700MS, T#2100MS, T#2400MS, T#1900MS, T#1700MS, T#1100MS, T#1700MS, T#2100MS, T#2900MS, T#2100MS, T#1700MS, T#1100MS, T#1700MS, T#1900MS, T#4800MS, T#2100MS, T#1700MS, T#1100MS, T#1700MS, T#2300MS, T#2300MS, T#1700MS, T#1100MS, T#1700MS, T#2100MS, T#2400MS, T#1900MS, T#1700MS, T#1100MS, T#1700MS, T#2100MS, T#1700MS, T#2100MS, T#1700MS, T#1100MS, T#1700MS, T#1900MS, T#3500MS, T#2100MS, T#1700MS, T#1100MS, T#1700MS, T#2300MS, T#2300MS, T#1700MS, T#1100MS, T#1700MS, T#2100MS, T#6000MS, T#1900MS, T#1700MS, T#1100MS, T#1700MS, T#2100MS, T#4100MS, T#2100MS, T#1700MS, T#1100MS, T#1700MS, T#1900MS, T#6000MS, T#2100MS, T#1700MS, T#1100MS, T#1700MS, T#2300MS, T#2300MS, T#1700MS, T#1100MS, T#1700MS, T#2100MS, T#2400MS, T#1900MS, T#1700MS, T#1100MS, T#1700MS, T#2100MS, T#4100MS, T#1100MS, T#1700MS, T#1100MS, T#1700MS, T#1100MS, T#6000MS, T#2100MS, T#1700MS, T#1100MS, T#1700MS, T#2300MS, T#2300MS, T#1700MS, T#1100MS, T#1700MS, T#2100MS, T#2400MS, T#1900MS, T#1700MS, T#1100MS, T#1700MS, T#2100MS, T#2900MS, T#1100MS, T#1700MS, T#1100MS, T#1700MS, T#1100MS, T#4800MS, T#2100MS, T#1700MS, T#1100MS, T#1700MS, T#2300MS, T#2300MS, T#1700MS, T#1100MS, T#1700MS, T#2100MS, T#2400MS, T#1900MS, T#1700MS, T#1100MS, T#1700MS, T#2100MS, T#1700MS, T#1100MS, T#1700MS, T#1100MS, T#1700MS, T#1100MS, T#3500MS, T#2100MS, T#1700MS, T#1100MS, T#1700MS, T#2300MS, T#2300MS, T#1700MS, T#1100MS, T#1700MS, T#2100MS, T#2400MS, T#1900MS, T#1700MS, T#1100MS, T#1700MS, T#2100MS, T#600MS, T#1100MS, T#1700MS, T#1100MS, T#1700MS, T#1100MS, T#2400MS, T#2100MS, T#1700MS, T#1100MS, T#1700MS, T#2300MS, T#2300MS, T#1700MS, T#1100MS, T#1700MS, T#2100MS, T#2400MS, T#1900MS, T#1700MS, T#1100MS, T#1700MS, T#2100MS, T#4100MS, T#1300MS, T#1700MS, T#1100MS, T#1700MS, T#1500MS, T#6000MS, T#2100MS, T#1700MS, T#1100MS, T#1700MS, T#2300MS, T#2300MS, T#1700MS, T#1100MS, T#1700MS, T#2100MS, T#2400MS, T#1900MS, T#1700MS, T#1100MS, T#1700MS, T#2100MS, T#2900MS, T#1300MS, T#1700MS, T#1100MS, T#1700MS, T#1500MS, T#4800MS, T#2100MS, T#1700MS, T#1100MS, T#1700MS, T#2300MS, T#2300MS, T#1700MS, T#1100MS, T#1700MS, T#2100MS, T#2400MS, T#1900MS, T#1700MS, T#1100MS, T#1700MS, T#2100MS, T#1700MS, T#1300MS, T#1700MS, T#1100MS, T#1700MS, T#1500MS, T#3500MS, T#2100MS, T#1700MS, T#1100MS, T#1700MS, T#2300MS, T#2300MS, T#1700MS, T#1100MS, T#1700MS, T#2100MS, T#2400MS, T#1900MS, T#1700MS, T#1100MS, T#1700MS, T#2100MS, T#600MS, T#1300MS, T#1700MS, T#1100MS, T#1700MS, T#1500MS, T#2400MS, T#2100MS, T#1700MS, T#1100MS, T#1700MS, T#2300MS, T#2300MS, T#1700MS, T#1100MS, T#1700MS, T#2100MS, T#6000MS, T#1100MS, T#1700MS, T#1100MS, T#1700MS, T#1100MS, T#600MS, T#2100MS, T#1700MS, T#1100MS, T#1700MS, T#1900MS, T#6000MS, T#2100MS, T#1700MS, T#1100MS, T#1700MS, T#2300MS, T#2300MS, T#1700MS, T#1100MS, T#1700MS, T#2100MS, T#6000MS, T#1100MS, T#1700MS, T#1100MS, T#1700MS, T#1100MS, T#1700MS, T#2100MS, T#1700MS, T#1100MS, T#1700MS, T#1900MS, T#4800MS, T#2100MS, T#1700MS, T#1100MS, T#1700MS, T#2300MS, T#2300MS, T#1700MS, T#1100MS, T#1700MS, T#2100MS, T#6000MS, T#1100MS, T#1700MS, T#1100MS, T#1700MS, T#1100MS, T#2900MS, T#2100MS, T#1700MS, T#1100MS, T#1700MS, T#1900MS, T#3500MS, T#2100MS, T#1700MS, T#1100MS, T#1700MS, T#2300MS, T#2300MS, T#1700MS, T#1100MS, T#1700MS, T#2100MS, T#6000MS, T#1100MS, T#1700MS, T#1100MS, T#1700MS, T#1100MS, T#4100MS, T#2100MS, T#1700MS, T#1100MS, T#1700MS, T#1900MS, T#2400MS, T#2100MS, T#1700MS, T#1100MS, T#1700MS, T#2300MS, T#2300MS, T#1700MS, T#1100MS, T#1700MS, T#2100MS, T#6000MS, T#1900MS, T#1700MS, T#1100MS, T#1700MS, T#2100MS, T#4100MS, T#2100MS, T#1700MS, T#1100MS, T#1700MS, T#1900MS, T#6000MS, T#2100MS, T#1700MS, T#1100MS, T#1700MS, T#2300MS, T#2300MS, T#1700MS, T#1100MS, T#1700MS, T#2100MS, T#6000MS, T#1100MS, T#1700MS, T#1100MS, T#1700MS, T#1100MS, T#1700MS, T#1100MS, T#1700MS, T#1100MS, T#1700MS, T#1100MS, T#4800MS, T#2100MS, T#1700MS, T#1100MS, T#1700MS, T#2300MS, T#2300MS, T#1700MS, T#1100MS, T#1700MS, T#2100MS, T#6000MS, T#1100MS, T#1700MS, T#1100MS, T#1700MS, T#1100MS, T#2900MS, T#1100MS, T#1700MS, T#1100MS, T#1700MS, T#1100MS, T#3500MS, T#2100MS, T#1700MS, T#1100MS, T#1700MS, T#2300MS, T#2300MS, T#1700MS, T#1100MS, T#1700MS, T#2100MS, T#6000MS, T#1100MS, T#1700MS, T#1100MS, T#1700MS, T#1100MS, T#4100MS, T#1100MS, T#1700MS, T#1100MS, T#1700MS, T#1100MS, T#2400MS, T#2100MS, T#1700MS, T#1100MS, T#1700MS, T#2300MS, T#2300MS, T#1700MS, T#1100MS, T#1700MS, T#2100MS, T#6000MS, T#1100MS, T#1700MS, T#1100MS, T#1700MS, T#1100MS, T#600MS, T#1300MS, T#1700MS, T#1100MS, T#1700MS, T#1500MS, T#6000MS, T#2100MS, T#1700MS, T#1100MS, T#1700MS, T#2300MS, T#2300MS, T#1700MS, T#1100MS, T#1700MS, T#2100MS, T#6000MS, T#1100MS, T#1700MS, T#1100MS, T#1700MS, T#1100MS, T#1700MS, T#1300MS, T#1700MS, T#1100MS, T#1700MS, T#1500MS, T#4800MS, T#2100MS, T#1700MS, T#1100MS, T#1700MS, T#2300MS, T#2300MS, T#1700MS, T#1100MS, T#1700MS, T#2100MS, T#6000MS, T#1100MS, T#1700MS, T#1100MS, T#1700MS, T#1100MS, T#2900MS, T#1300MS, T#1700MS, T#1100MS, T#1700MS, T#1500MS, T#3500MS, T#2100MS, T#1700MS, T#1100MS, T#1700MS, T#2300MS, T#2300MS, T#1700MS, T#1100MS, T#1700MS, T#2100MS, T#6000MS, T#1100MS, T#1700MS, T#1100MS, T#1700MS, T#1100MS, T#4100MS, T#1300MS, T#1700MS, T#1100MS, T#1700MS, T#1500MS, T#2400MS, T#2100MS, T#1700MS, T#1100MS, T#1700MS, T#2300MS, T#2300MS, T#1700MS, T#1100MS, T#1700MS, T#2100MS, T#4800MS, T#1100MS, T#1700MS, T#1100MS, T#1700MS, T#1100MS, T#1700MS, T#2100MS, T#1700MS, T#1100MS, T#1700MS, T#1900MS, T#6000MS, T#2100MS, T#1700MS, T#1100MS, T#1700MS, T#2300MS, T#2300MS, T#1700MS, T#1100MS, T#1700MS, T#2100MS, T#4800MS, T#1100MS, T#1700MS, T#1100MS, T#1700MS, T#1100MS, T#600MS, T#2100MS, T#1700MS, T#1100MS, T#1700MS, T#1900MS, T#4800MS, T#2100MS, T#1700MS, T#1100MS, T#1700MS, T#2300MS, T#2300MS, T#1700MS, T#1100MS, T#1700MS, T#2100MS, T#4800MS, T#1100MS, T#1700MS, T#1100MS, T#1700MS, T#1100MS, T#1700MS, T#2100MS, T#1700MS, T#1100MS, T#1700MS, T#1900MS, T#3500MS, T#2100MS, T#1700MS, T#1100MS, T#1700MS, T#2300MS, T#2300MS, T#1700MS, T#1100MS, T#1700MS, T#2100MS, T#4800MS, T#1100MS, T#1700MS, T#1100MS, T#1700MS, T#1100MS, T#2900MS, T#2100MS, T#1700MS, T#1100MS, T#1700MS, T#1900MS, T#2400MS, T#2100MS, T#1700MS, T#1100MS, T#1700MS, T#2300MS, T#2300MS, T#1700MS, T#1100MS, T#1700MS, T#2100MS, T#4800MS, T#1100MS, T#1700MS, T#1100MS, T#1700MS, T#1100MS, T#1700MS, T#1100MS, T#1700MS, T#1100MS, T#1700MS, T#1100MS, T#6000MS, T#2100MS, T#1700MS, T#1100MS, T#1700MS, T#2300MS, T#2300MS, T#1700MS, T#1100MS, T#1700MS, T#2100MS, T#6000MS, T#1900MS, T#1700MS, T#1100MS, T#1700MS, T#2100MS, T#4100MS, T#2100MS, T#1700MS, T#1100MS, T#1700MS, T#1900MS, T#6000MS, T#2100MS, T#1700MS, T#1100MS, T#1700MS, T#2300MS, T#2300MS, T#1700MS, T#1100MS, T#1700MS, T#2100MS, T#4800MS, T#1100MS, T#1700MS, T#1100MS, T#1700MS, T#1100MS, T#1700MS, T#1100MS, T#1700MS, T#1100MS, T#1700MS, T#1100MS, T#3500MS, T#2100MS, T#1700MS, T#1100MS, T#1700MS, T#2300MS, T#2300MS, T#1700MS, T#1100MS, T#1700MS, T#2100MS, T#4800MS, T#1100MS, T#1700MS, T#1100MS, T#1700MS, T#1100MS, T#2900MS, T#1100MS, T#1700MS, T#1100MS, T#1700MS, T#1100MS, T#2400MS, T#2100MS, T#1700MS, T#1100MS, T#1700MS, T#2300MS, T#2300MS, T#1700MS, T#1100MS, T#1700MS, T#2100MS, T#4800MS, T#1100MS, T#1700MS, T#1100MS, T#1700MS, T#1100MS, T#1700MS, T#1300MS, T#1700MS, T#1100MS, T#1700MS, T#1500MS, T#6000MS, T#2100MS, T#1700MS, T#1100MS, T#1700MS, T#2300MS, T#2300MS, T#1700MS, T#1100MS, T#1700MS, T#2100MS, T#4800MS, T#1100MS, T#1700MS, T#1100MS, T#1700MS, T#1100MS, T#600MS, T#1300MS, T#1700MS, T#1100MS, T#1700MS, T#1500MS, T#4800MS, T#2100MS, T#1700MS, T#1100MS, T#1700MS, T#2300MS, T#2300MS, T#1700MS, T#1100MS, T#1700MS, T#2100MS, T#4800MS, T#1100MS, T#1700MS, T#1100MS, T#1700MS, T#1100MS, T#1700MS, T#1300MS, T#1700MS, T#1100MS, T#1700MS, T#1500MS, T#3500MS, T#2100MS, T#1700MS, T#1100MS, T#1700MS, T#2300MS, T#2300MS, T#1700MS, T#1100MS, T#1700MS, T#2100MS, T#4800MS, T#1100MS, T#1700MS, T#1100MS, T#1700MS, T#1100MS, T#2900MS, T#1300MS, T#1700MS, T#1100MS, T#1700MS, T#1500MS, T#2400MS, T#2100MS, T#1700MS, T#1100MS, T#1700MS, T#2300MS, T#2300MS, T#1700MS, T#1100MS, T#1700MS, T#2100MS, T#3500MS, T#1100MS, T#1700MS, T#1100MS, T#1700MS, T#1100MS, T#2900MS, T#2100MS, T#1700MS, T#1100MS, T#1700MS, T#1900MS, T#6000MS, T#2100MS, T#1700MS, T#1100MS, T#1700MS, T#2300MS, T#2300MS, T#1700MS, T#1100MS, T#1700MS, T#2100MS, T#3500MS, T#1100MS, T#1700MS, T#1100MS, T#1700MS, T#1100MS, T#1700MS, T#2100MS, T#1700MS, T#1100MS, T#1700MS, T#1900MS, T#4800MS, T#2100MS, T#1700MS, T#1100MS, T#1700MS, T#2300MS, T#2300MS, T#1700MS, T#1100MS, T#1700MS, T#2100MS, T#3500MS, T#1100MS, T#1700MS, T#1100MS, T#1700MS, T#1100MS, T#600MS, T#2100MS, T#1700MS, T#1100MS, T#1700MS, T#1900MS, T#3500MS, T#2100MS, T#1700MS, T#1100MS, T#1700MS, T#2300MS, T#2300MS, T#1700MS, T#1100MS, T#1700MS, T#2100MS, T#3500MS, T#1100MS, T#1700MS, T#1100MS, T#1700MS, T#1100MS, T#1700MS, T#2100MS, T#1700MS, T#1100MS, T#1700MS, T#1900MS, T#2400MS, T#2100MS, T#1700MS, T#1100MS, T#1700MS, T#2300MS, T#2300MS, T#1700MS, T#1100MS, T#1700MS, T#2100MS, T#3500MS, T#1100MS, T#1700MS, T#1100MS, T#1700MS, T#1100MS, T#2900MS, T#1100MS, T#1700MS, T#1100MS, T#1700MS, T#1100MS, T#6000MS, T#2100MS, T#1700MS, T#1100MS, T#1700MS, T#2300MS, T#2300MS, T#1700MS, T#1100MS, T#1700MS, T#2100MS, T#3500MS, T#1100MS, T#1700MS, T#1100MS, T#1700MS, T#1100MS, T#1700MS, T#1100MS, T#1700MS, T#1100MS, T#1700MS, T#1100MS, T#4800MS, T#2100MS, T#1700MS, T#1100MS, T#1700MS, T#2300MS, T#2300MS, T#1700MS, T#1100MS, T#1700MS, T#2100MS, T#6000MS, T#1900MS, T#1700MS, T#1100MS, T#1700MS, T#2100MS, T#4100MS, T#2100MS, T#1700MS, T#1100MS, T#1700MS, T#1900MS, T#6000MS, T#2100MS, T#1700MS, T#1100MS, T#1700MS, T#2300MS, T#2300MS, T#1700MS, T#1100MS, T#1700MS, T#2100MS, T#3500MS, T#1100MS, T#1700MS, T#1100MS, T#1700MS, T#1100MS, T#1700MS, T#1100MS, T#1700MS, T#1100MS, T#1700MS, T#1100MS, T#2400MS, T#2100MS, T#1700MS, T#1100MS, T#1700MS, T#2300MS, T#2300MS, T#1700MS, T#1100MS, T#1700MS, T#2100MS, T#3500MS, T#1100MS, T#1700MS, T#1100MS, T#1700MS, T#1100MS, T#2900MS, T#1300MS, T#1700MS, T#1100MS, T#1700MS, T#1500MS, T#6000MS, T#2100MS, T#1700MS, T#1100MS, T#1700MS, T#2300MS, T#2300MS, T#1700MS, T#1100MS, T#1700MS, T#2100MS, T#3500MS, T#1100MS, T#1700MS, T#1100MS, T#1700MS, T#1100MS, T#1700MS, T#1300MS, T#1700MS, T#1100MS, T#1700MS, T#1500MS, T#4800MS, T#2100MS, T#1700MS, T#1100MS, T#1700MS, T#2300MS, T#2300MS, T#1700MS, T#1100MS, T#1700MS, T#2100MS, T#3500MS, T#1100MS, T#1700MS, T#1100MS, T#1700MS, T#1100MS, T#600MS, T#1300MS, T#1700MS, T#1100MS, T#1700MS, T#1500MS, T#3500MS, T#2100MS, T#1700MS, T#1100MS, T#1700MS, T#2300MS, T#2300MS, T#1700MS, T#1100MS, T#1700MS, T#2100MS, T#3500MS, T#1100MS, T#1700MS, T#1100MS, T#1700MS, T#1100MS, T#1700MS, T#1300MS, T#1700MS, T#1100MS, T#1700MS, T#1500MS, T#2400MS, T#2100MS, T#1700MS, T#1100MS, T#1700MS, T#2300MS, T#2300MS, T#1700MS, T#1100MS, T#1700MS, T#2100MS, T#2400MS, T#1100MS, T#1700MS, T#1100MS, T#1700MS, T#1100MS, T#4100MS, T#2100MS, T#1700MS, T#1100MS, T#1700MS, T#1900MS, T#6000MS, T#2100MS, T#1700MS, T#1100MS, T#1700MS, T#2300MS, T#2300MS, T#1700MS, T#1100MS, T#1700MS, T#2100MS, T#2400MS, T#1100MS, T#1700MS, T#1100MS, T#1700MS, T#1100MS, T#2900MS, T#2100MS, T#1700MS, T#1100MS, T#1700MS, T#1900MS, T#4800MS, T#2100MS, T#1700MS, T#1100MS, T#1700MS, T#2300MS, T#2300MS, T#1700MS, T#1100MS, T#1700MS, T#2100MS, T#2400MS, T#1100MS, T#1700MS, T#1100MS, T#1700MS, T#1100MS, T#1700MS, T#2100MS, T#1700MS, T#1100MS, T#1700MS, T#1900MS, T#3500MS, T#2100MS, T#1700MS, T#1100MS, T#1700MS, T#2300MS, T#2300MS, T#1700MS, T#1100MS, T#1700MS, T#2100MS, T#2400MS, T#1100MS, T#1700MS, T#1100MS, T#1700MS, T#1100MS, T#600MS, T#2100MS, T#1700MS, T#1100MS, T#1700MS, T#1900MS, T#2400MS, T#2100MS, T#1700MS, T#1100MS, T#1700MS, T#2300MS, T#2300MS, T#1700MS, T#1100MS, T#1700MS, T#2100MS, T#2400MS, T#1100MS, T#1700MS, T#1100MS, T#1700MS, T#1100MS, T#4100MS, T#1100MS, T#1700MS, T#1100MS, T#1700MS, T#1100MS, T#6000MS, T#2100MS, T#1700MS, T#1100MS, T#1700MS, T#2300MS, T#2300MS, T#1700MS, T#1100MS, T#1700MS, T#2100MS, T#2400MS, T#1100MS, T#1700MS, T#1100MS, T#1700MS, T#1100MS, T#2900MS, T#1100MS, T#1700MS, T#1100MS, T#1700MS, T#1100MS, T#4800MS, T#2100MS, T#1700MS, T#1100MS, T#1700MS, T#2300MS, T#2300MS, T#1700MS, T#1100MS, T#1700MS, T#2100MS, T#2400MS, T#1100MS, T#1700MS, T#1100MS, T#1700MS, T#1100MS, T#1700MS, T#1100MS, T#1700MS, T#1100MS, T#1700MS, T#1100MS, T#3500MS, T#2100MS, T#1700MS, T#1100MS, T#1700MS, T#2300MS, T#2300MS, T#1700MS, T#1100MS, T#1700MS, T#2100MS, T#6000MS, T#1900MS, T#1700MS, T#1100MS, T#1700MS, T#2100MS, T#4100MS, T#2100MS, T#1700MS, T#1100MS, T#1700MS, T#1900MS, T#6000MS, T#2100MS, T#1700MS, T#1100MS, T#1700MS, T#2300MS, T#2300MS, T#1700MS, T#1100MS, T#1700MS, T#2100MS, T#2400MS, T#1100MS, T#1700MS, T#1100MS, T#1700MS, T#1100MS, T#4100MS, T#1300MS, T#1700MS, T#1100MS, T#1700MS, T#1500MS, T#6000MS, T#2100MS, T#1700MS, T#1100MS, T#1700MS, T#2300MS, T#2300MS, T#1700MS, T#1100MS, T#1700MS, T#2100MS, T#2400MS, T#1100MS, T#1700MS, T#1100MS, T#1700MS, T#1100MS, T#2900MS, T#1300MS, T#1700MS, T#1100MS, T#1700MS, T#1500MS, T#4800MS, T#2100MS, T#1700MS, T#1100MS, T#1700MS, T#2300MS, T#2300MS, T#1700MS, T#1100MS, T#1700MS, T#2100MS, T#2400MS, T#1100MS, T#1700MS, T#1100MS, T#1700MS, T#1100MS, T#1700MS, T#1300MS, T#1700MS, T#1100MS, T#1700MS, T#1500MS, T#3500MS, T#2100MS, T#1700MS, T#1100MS, T#1700MS, T#2300MS, T#2300MS, T#1700MS, T#1100MS, T#1700MS, T#2100MS, T#2400MS, T#1100MS, T#1700MS, T#1100MS, T#1700MS, T#1100MS, T#600MS, T#1300MS, T#1700MS, T#1100MS, T#1700MS, T#1500MS, T#2400MS, T#2100MS, T#1700MS, T#1100MS, T#1700MS, T#2300MS, T#2300MS, T#1700MS, T#1100MS, T#1700MS, T#2100MS, T#6000MS, T#1500MS, T#1700MS, T#1100MS, T#1700MS, T#1300MS, T#600MS, T#2100MS, T#1700MS, T#1100MS, T#1700MS, T#1900MS, T#6000MS, T#2100MS, T#1700MS, T#1100MS, T#1700MS, T#2300MS, T#2300MS, T#1700MS, T#1100MS, T#1700MS, T#2100MS, T#6000MS, T#1500MS, T#1700MS, T#1100MS, T#1700MS, T#1300MS, T#1700MS, T#2100MS, T#1700MS, T#1100MS, T#1700MS, T#1900MS, T#4800MS, T#2100MS, T#1700MS, T#1100MS, T#1700MS, T#2300MS, T#2300MS, T#1700MS, T#1100MS, T#1700MS, T#2100MS, T#6000MS, T#1500MS, T#1700MS, T#1100MS, T#1700MS, T#1300MS, T#2900MS, T#2100MS, T#1700MS, T#1100MS, T#1700MS, T#1900MS, T#3500MS, T#2100MS, T#1700MS, T#1100MS, T#1700MS, T#2300MS, T#2300MS, T#1700MS, T#1100MS, T#1700MS, T#2100MS, T#6000MS, T#1500MS, T#1700MS, T#1100MS, T#1700MS, T#1300MS, T#4100MS, T#2100MS, T#1700MS, T#1100MS, T#1700MS, T#1900MS, T#2400MS, T#2100MS, T#1700MS, T#1100MS, T#1700MS, T#2300MS, T#2300MS, T#1700MS, T#1100MS, T#1700MS, T#2100MS, T#6000MS, T#1500MS, T#1700MS, T#1100MS, T#1700MS, T#1300MS, T#600MS, T#1100MS, T#1700MS, T#1100MS, T#1700MS, T#1100MS, T#6000MS, T#2100MS, T#1700MS, T#1100MS, T#1700MS, T#2300MS, T#2300MS, T#1700MS, T#1100MS, T#1700MS, T#2100MS, T#6000MS, T#1500MS, T#1700MS, T#1100MS, T#1700MS, T#1300MS, T#1700MS, T#1100MS, T#1700MS, T#1100MS, T#1700MS, T#1100MS, T#4800MS, T#2100MS, T#1700MS, T#1100MS, T#1700MS, T#2300MS, T#2300MS, T#1700MS, T#1100MS, T#1700MS, T#2100MS, T#6000MS, T#1500MS, T#1700MS, T#1100MS, T#1700MS, T#1300MS, T#2900MS, T#1100MS, T#1700MS, T#1100MS, T#1700MS, T#1100MS, T#3500MS, T#2100MS, T#1700MS, T#1100MS, T#1700MS, T#2300MS, T#2300MS, T#1700MS, T#1100MS, T#1700MS, T#2100MS, T#6000MS, T#1500MS, T#1700MS, T#1100MS, T#1700MS, T#1300MS, T#4100MS, T#1100MS, T#1700MS, T#1100MS, T#1700MS, T#1100MS, T#2400MS, T#2100MS, T#1700MS, T#1100MS, T#1700MS, T#2300MS, T#2300MS, T#1700MS, T#1100MS, T#1700MS, T#2100MS, T#6000MS, T#1900MS, T#1700MS, T#1100MS, T#1700MS, T#2100MS, T#4100MS, T#2100MS, T#1700MS, T#1100MS, T#1700MS, T#1900MS, T#6000MS, T#2100MS, T#1700MS, T#1100MS, T#1700MS, T#2300MS, T#2300MS, T#1700MS, T#1100MS, T#1700MS, T#2100MS, T#6000MS, T#1500MS, T#1700MS, T#1100MS, T#1700MS, T#1300MS, T#1700MS, T#1300MS, T#1700MS, T#1100MS, T#1700MS, T#1500MS, T#4800MS, T#2100MS, T#1700MS, T#1100MS, T#1700MS, T#2300MS, T#2300MS, T#1700MS, T#1100MS, T#1700MS, T#2100MS, T#6000MS, T#1500MS, T#1700MS, T#1100MS, T#1700MS, T#1300MS, T#2900MS, T#1300MS, T#1700MS, T#1100MS, T#1700MS, T#1500MS, T#3500MS, T#2100MS, T#1700MS, T#1100MS, T#1700MS, T#2300MS, T#2300MS, T#1700MS, T#1100MS, T#1700MS, T#2100MS, T#6000MS, T#1500MS, T#1700MS, T#1100MS, T#1700MS, T#1300MS, T#4100MS, T#1300MS, T#1700MS, T#1100MS, T#1700MS, T#1500MS, T#2400MS, T#2100MS, T#1700MS, T#1100MS, T#1700MS, T#2300MS, T#2300MS, T#1700MS, T#1100MS, T#1700MS, T#2100MS, T#4800MS, T#1500MS, T#1700MS, T#1100MS, T#1700MS, T#1300MS, T#1700MS, T#2100MS, T#1700MS, T#1100MS, T#1700MS, T#1900MS, T#6000MS, T#2100MS, T#1700MS, T#1100MS, T#1700MS, T#2300MS, T#2300MS, T#1700MS, T#1100MS, T#1700MS, T#2100MS, T#4800MS, T#1500MS, T#1700MS, T#1100MS, T#1700MS, T#1300MS, T#600MS, T#2100MS, T#1700MS, T#1100MS, T#1700MS, T#1900MS, T#4800MS, T#2100MS, T#1700MS, T#1100MS, T#1700MS, T#2300MS, T#2300MS, T#1700MS, T#1100MS, T#1700MS, T#2100MS, T#4800MS, T#1500MS, T#1700MS, T#1100MS, T#1700MS, T#1300MS, T#1700MS, T#2100MS, T#1700MS, T#1100MS, T#1700MS, T#1900MS, T#3500MS, T#2100MS, T#1700MS, T#1100MS, T#1700MS, T#2300MS, T#2300MS, T#1700MS, T#1100MS, T#1700MS, T#2100MS, T#4800MS, T#1500MS, T#1700MS, T#1100MS, T#1700MS, T#1300MS, T#2900MS, T#2100MS, T#1700MS, T#1100MS, T#1700MS, T#1900MS, T#2400MS, T#2100MS, T#1700MS, T#1100MS, T#1700MS, T#2300MS, T#2300MS, T#1700MS, T#1100MS, T#1700MS, T#2100MS, T#4800MS, T#1500MS, T#1700MS, T#1100MS, T#1700MS, T#1300MS, T#1700MS, T#1100MS, T#1700MS, T#1100MS, T#1700MS, T#1100MS, T#6000MS, T#2100MS, T#1700MS, T#1100MS, T#1700MS, T#2300MS, T#2300MS, T#1700MS, T#1100MS, T#1700MS, T#2100MS, T#4800MS, T#1500MS, T#1700MS, T#1100MS, T#1700MS, T#1300MS, T#600MS, T#1100MS, T#1700MS, T#1100MS, T#1700MS, T#1100MS, T#4800MS, T#2100MS, T#1700MS, T#1100MS, T#1700MS, T#2300MS, T#2300MS, T#1700MS, T#1100MS, T#1700MS, T#2100MS, T#4800MS, T#1500MS, T#1700MS, T#1100MS, T#1700MS, T#1300MS, T#1700MS, T#1100MS, T#1700MS, T#1100MS, T#1700MS, T#1100MS, T#3500MS, T#2100MS, T#1700MS, T#1100MS, T#1700MS, T#2300MS, T#2300MS, T#1700MS, T#1100MS, T#1700MS, T#2100MS, T#4800MS, T#1500MS, T#1700MS, T#1100MS, T#1700MS, T#1300MS, T#2900MS, T#1100MS, T#1700MS, T#1100MS, T#1700MS, T#1100MS, T#2400MS, T#2100MS, T#1700MS, T#1100MS, T#1700MS, T#2300MS, T#2300MS, T#1700MS, T#1100MS, T#1700MS, T#2100MS, T#4800MS, T#1500MS, T#1700MS, T#1100MS, T#1700MS, T#1300MS, T#1700MS, T#1300MS, T#1700MS, T#1100MS, T#1700MS, T#1500MS, T#6000MS, T#2100MS, T#1700MS, T#1100MS, T#1700MS, T#2300MS, T#2300MS, T#1700MS, T#1100MS, T#1700MS, T#2100MS, T#6000MS, T#1900MS, T#1700MS, T#1100MS, T#1700MS, T#2100MS, T#4100MS, T#2100MS, T#1700MS, T#1100MS, T#1700MS, T#1900MS, T#6000MS, T#2100MS, T#1700MS, T#1100MS, T#1700MS, T#2300MS, T#2300MS, T#1700MS, T#1100MS, T#1700MS, T#2100MS, T#4800MS, T#1500MS, T#1700MS, T#1100MS, T#1700MS, T#1300MS, T#1700MS, T#1300MS, T#1700MS, T#1100MS, T#1700MS, T#1500MS, T#3500MS, T#2100MS, T#1700MS, T#1100MS, T#1700MS, T#2300MS, T#2300MS, T#1700MS, T#1100MS, T#1700MS, T#2100MS, T#4800MS, T#1500MS, T#1700MS, T#1100MS, T#1700MS, T#1300MS, T#2900MS, T#1300MS, T#1700MS, T#1100MS, T#1700MS, T#1500MS, T#2400MS, T#2100MS, T#1700MS, T#1100MS, T#1700MS, T#2300MS, T#2300MS, T#1700MS, T#1100MS, T#1700MS, T#2100MS, T#3500MS, T#1500MS, T#1700MS, T#1100MS, T#1700MS, T#1300MS, T#2900MS, T#2100MS, T#1700MS, T#1100MS, T#1700MS, T#1900MS, T#6000MS, T#2100MS, T#1700MS, T#1100MS, T#1700MS, T#2300MS, T#2300MS, T#1700MS, T#1100MS, T#1700MS, T#2100MS, T#3500MS, T#1500MS, T#1700MS, T#1100MS, T#1700MS, T#1300MS, T#1700MS, T#2100MS, T#1700MS, T#1100MS, T#1700MS, T#1900MS, T#4800MS, T#2100MS, T#1700MS, T#1100MS, T#1700MS, T#2300MS, T#2300MS, T#1700MS, T#1100MS, T#1700MS, T#2100MS, T#3500MS, T#1500MS, T#1700MS, T#1100MS, T#1700MS, T#1300MS, T#600MS, T#2100MS, T#1700MS, T#1100MS, T#1700MS, T#1900MS, T#3500MS, T#2100MS, T#1700MS, T#1100MS, T#1700MS, T#2300MS, T#2300MS, T#1700MS, T#1100MS, T#1700MS, T#2100MS, T#3500MS, T#1500MS, T#1700MS, T#1100MS, T#1700MS, T#1300MS, T#1700MS, T#2100MS, T#1700MS, T#1100MS, T#1700MS, T#1900MS, T#2400MS, T#2100MS, T#1700MS, T#1100MS, T#1700MS, T#2300MS, T#2300MS, T#1700MS, T#1100MS, T#1700MS, T#2100MS, T#3500MS, T#1500MS, T#1700MS, T#1100MS, T#1700MS, T#1300MS, T#2900MS, T#1100MS, T#1700MS, T#1100MS, T#1700MS, T#1100MS, T#6000MS, T#2100MS, T#1700MS, T#1100MS, T#1700MS, T#2300MS, T#2300MS, T#1700MS, T#1100MS, T#1700MS, T#2100MS, T#3500MS, T#1500MS, T#1700MS, T#1100MS, T#1700MS, T#1300MS, T#1700MS, T#1100MS, T#1700MS, T#1100MS, T#1700MS, T#1100MS, T#4800MS, T#2100MS, T#1700MS, T#1100MS, T#1700MS, T#2300MS, T#2300MS, T#1700MS, T#1100MS, T#1700MS, T#2100MS, T#3500MS, T#1500MS, T#1700MS, T#1100MS, T#1700MS, T#1300MS, T#600MS, T#1100MS, T#1700MS, T#1100MS, T#1700MS, T#1100MS, T#3500MS, T#2100MS, T#1700MS, T#1100MS, T#1700MS, T#2300MS, T#2300MS, T#1700MS, T#1100MS, T#1700MS, T#2100MS, T#3500MS, T#1500MS, T#1700MS, T#1100MS, T#1700MS, T#1300MS, T#1700MS, T#1100MS, T#1700MS, T#1100MS, T#1700MS, T#1100MS, T#2400MS, T#2100MS, T#1700MS, T#1100MS, T#1700MS, T#2300MS, T#2300MS, T#1700MS, T#1100MS, T#1700MS, T#2100MS, T#3500MS, T#1500MS, T#1700MS, T#1100MS, T#1700MS, T#1300MS, T#2900MS, T#1300MS, T#1700MS, T#1100MS, T#1700MS, T#1500MS, T#6000MS, T#2100MS, T#1700MS, T#1100MS, T#1700MS, T#2300MS, T#2300MS, T#1700MS, T#1100MS, T#1700MS, T#2100MS, T#3500MS, T#1500MS, T#1700MS, T#1100MS, T#1700MS, T#1300MS, T#1700MS, T#1300MS, T#1700MS, T#1100MS, T#1700MS, T#1500MS, T#4800MS, T#2100MS, T#1700MS, T#1100MS, T#1700MS, T#2300MS, T#2300MS, T#1700MS, T#1100MS, T#1700MS, T#2100MS, T#6000MS, T#1900MS, T#1700MS, T#1100MS, T#1700MS, T#2100MS, T#4100MS, T#2100MS, T#1700MS, T#1100MS, T#1700MS, T#1900MS, T#6000MS, T#2100MS, T#1700MS, T#1100MS, T#1700MS, T#2300MS, T#2300MS, T#1700MS, T#1100MS, T#1700MS, T#2100MS, T#3500MS, T#1500MS, T#1700MS, T#1100MS, T#1700MS, T#1300MS, T#1700MS, T#1300MS, T#1700MS, T#1100MS, T#1700MS, T#1500MS, T#2400MS, T#2100MS, T#1700MS, T#1100MS, T#1700MS, T#2300MS, T#2300MS, T#1700MS, T#1100MS, T#1700MS, T#2100MS, T#2400MS, T#1500MS, T#1700MS, T#1100MS, T#1700MS, T#1300MS, T#4100MS, T#2100MS, T#1700MS, T#1100MS, T#1700MS, T#1900MS, T#6000MS, T#2100MS, T#1700MS, T#1100MS, T#1700MS, T#2300MS, T#2300MS, T#1700MS, T#1100MS, T#1700MS, T#2100MS, T#2400MS, T#1500MS, T#1700MS, T#1100MS, T#1700MS, T#1300MS, T#2900MS, T#2100MS, T#1700MS, T#1100MS, T#1700MS, T#1900MS, T#4800MS, T#2100MS, T#1700MS, T#1100MS, T#1700MS, T#2300MS, T#2300MS, T#1700MS, T#1100MS, T#1700MS, T#2100MS, T#2400MS, T#1500MS, T#1700MS, T#1100MS, T#1700MS, T#1300MS, T#1700MS, T#2100MS, T#1700MS, T#1100MS, T#1700MS, T#1900MS, T#3500MS, T#2100MS, T#1700MS, T#1100MS, T#1700MS, T#2300MS, T#2300MS, T#1700MS, T#1100MS, T#1700MS, T#2100MS, T#2400MS, T#1500MS, T#1700MS, T#1100MS, T#1700MS, T#1300MS, T#600MS, T#2100MS, T#1700MS, T#1100MS, T#1700MS, T#1900MS, T#2400MS, T#2100MS, T#1700MS, T#1100MS, T#1700MS, T#2300MS, T#2300MS, T#1700MS, T#1100MS, T#1700MS, T#2100MS, T#2400MS, T#1500MS, T#1700MS, T#1100MS, T#1700MS, T#1300MS, T#4100MS, T#1100MS, T#1700MS, T#1100MS, T#1700MS, T#1100MS, T#6000MS, T#2100MS, T#1700MS, T#1100MS, T#1700MS, T#2300MS, T#2300MS, T#1700MS, T#1100MS, T#1700MS, T#2100MS, T#2400MS, T#1500MS, T#1700MS, T#1100MS, T#1700MS, T#1300MS, T#2900MS, T#1100MS, T#1700MS, T#1100MS, T#1700MS, T#1100MS, T#4800MS, T#2100MS, T#1700MS, T#1100MS, T#1700MS, T#2300MS, T#2300MS, T#1700MS, T#1100MS, T#1700MS, T#2100MS, T#2400MS, T#1500MS, T#1700MS, T#1100MS, T#1700MS, T#1300MS, T#1700MS, T#1100MS, T#1700MS, T#1100MS, T#1700MS, T#1100MS, T#3500MS, T#2100MS, T#1700MS, T#1100MS, T#1700MS, T#2300MS, T#2300MS, T#1700MS, T#1100MS, T#1700MS, T#2100MS, T#2400MS, T#1500MS, T#1700MS, T#1100MS, T#1700MS, T#1300MS, T#600MS, T#1100MS, T#1700MS, T#1100MS, T#1700MS, T#1100MS, T#2400MS, T#2100MS, T#1700MS, T#1100MS, T#1700MS, T#2300MS, T#2300MS, T#1700MS, T#1100MS, T#1700MS, T#2100MS, T#2400MS, T#1500MS, T#1700MS, T#1100MS, T#1700MS, T#1300MS, T#4100MS, T#1300MS, T#1700MS, T#1100MS, T#1700MS, T#1500MS, T#6000MS, T#2100MS, T#1700MS, T#1100MS, T#1700MS, T#2300MS, T#2300MS, T#1700MS, T#1100MS, T#1700MS, T#2100MS, T#2400MS, T#1500MS, T#1700MS, T#1100MS, T#1700MS, T#1300MS, T#2900MS, T#1300MS, T#1700MS, T#1100MS, T#1700MS, T#1500MS, T#4800MS, T#2100MS, T#1700MS, T#1100MS, T#1700MS, T#2300MS, T#2300MS, T#1700MS, T#1100MS, T#1700MS, T#2100MS, T#2400MS, T#1500MS, T#1700MS, T#1100MS, T#1700MS, T#1300MS, T#1700MS, T#1300MS, T#1700MS, T#1100MS, T#1700MS, T#1500MS, T#3500MS, T#2100MS, T#1700MS, T#1100MS, T#1700MS, T#2300MS];
    WD_STORE : ARRAY[1..12, 1..12] OF TIME := [T#2300MS, T#1700MS, T#1100MS, T#1700MS, T#2100MS, T#6000MS, T#1900MS, T#1700MS, T#1100MS, T#1700MS, T#2100MS, T#6000MS, T#2300MS, T#1700MS, T#1100MS, T#1700MS, T#2100MS, T#4800MS, T#1900MS, T#1700MS, T#1100MS, T#1700MS, T#2100MS, T#4800MS, T#2300MS, T#1700MS, T#1100MS, T#1700MS, T#2100MS, T#3500MS, T#1900MS, T#1700MS, T#1100MS, T#1700MS, T#2100MS, T#3500MS, T#2300MS, T#1700MS, T#1100MS, T#1700MS, T#2100MS, T#2400MS, T#1900MS, T#1700MS, T#1100MS, T#1700MS, T#2100MS, T#2400MS, T#2300MS, T#1700MS, T#1100MS, T#1700MS, T#2100MS, T#6000MS, T#1100MS, T#1700MS, T#1100MS, T#1700MS, T#1100MS, T#6000MS, T#2300MS, T#1700MS, T#1100MS, T#1700MS, T#2100MS, T#4800MS, T#1100MS, T#1700MS, T#1100MS, T#1700MS, T#1100MS, T#4800MS, T#2300MS, T#1700MS, T#1100MS, T#1700MS, T#2100MS, T#3500MS, T#1100MS, T#1700MS, T#1100MS, T#1700MS, T#1100MS, T#3500MS, T#2300MS, T#1700MS, T#1100MS, T#1700MS, T#2100MS, T#2400MS, T#1100MS, T#1700MS, T#1100MS, T#1700MS, T#1100MS, T#2400MS, T#2300MS, T#1700MS, T#1100MS, T#1700MS, T#2100MS, T#6000MS, T#1500MS, T#1700MS, T#1100MS, T#1700MS, T#1300MS, T#6000MS, T#2300MS, T#1700MS, T#1100MS, T#1700MS, T#2100MS, T#4800MS, T#1500MS, T#1700MS, T#1100MS, T#1700MS, T#1300MS, T#4800MS, T#2300MS, T#1700MS, T#1100MS, T#1700MS, T#2100MS, T#3500MS, T#1500MS, T#1700MS, T#1100MS, T#1700MS, T#1300MS, T#3500MS, T#2300MS, T#1700MS, T#1100MS, T#1700MS, T#2100MS, T#2400MS, T#1500MS, T#1700MS, T#1100MS, T#1700MS, T#1300MS, T#2400MS];
    WD_FETCH_EMPTY : ARRAY[1..12, 1..12] OF TIME := [T#6000MS, T#2100MS, T#1700MS, T#1100MS, T#1700MS, T#1900MS, T#6000MS, T#2100MS, T#1700MS, T#1100MS, T#1700MS, T#2300MS, T#4800MS, T#2100MS, T#1700MS, T#1100MS, T#1700MS, T#1900MS, T#4800MS, T#2100MS, T#1700MS, T#1100MS, T#1700MS, T#2300MS, T#3500MS, T#2100MS, T#1700MS, T#1100MS, T#1700MS, T#1900MS, T#3500MS, T#2100MS, T#1700MS, T#1100MS, T#1700MS, T#2300MS, T#2400MS, T#2100MS, T#1700MS, T#1100MS, T#1700MS, T#1900MS, T#2400MS, T#2100MS, T#1700MS, T#1100MS, T#1700MS, T#2300MS, T#6000MS, T#1100MS, T#1700MS, T#1100MS, T#1700MS, T#1100MS, T#6000MS, T#2100MS, T#1700MS, T#1100MS, T#1700MS, T#2300MS, T#4800MS, T#1100MS, T#1700MS, T#1100MS, T#1700MS, T#1100MS, T#4800MS, T#2100MS, T#1700MS, T#1100MS, T#1700MS, T#2300MS, T#3500MS, T#1100MS, T#1700MS, T#1100MS, T#1700MS, T#1100MS, T#3500MS, T#2100MS, T#1700MS, T#1100MS, T#1700MS, T#2300MS, T#2400MS, T#1100MS, T#1700MS, T#1100MS, T#1700MS, T#1100MS, T#2400MS, T#2100MS, T#1700MS, T#1100MS, T#1700MS, T#2300MS, T#6000MS, T#1300MS, T#1700MS, T#1100MS, T#1700MS, T#1500MS, T#6000MS, T#2100MS, T#1700MS, T#1100MS, T#1700MS, T#2300MS, T#4800MS, T#1300MS, T#1700MS, T#1100MS, T#1700MS, T#1500MS, T#4800MS, T#2100MS, T#1700MS, T#1100MS, T#1700MS, T#2300MS, T#3500MS, T#1300MS, T#1700MS, T#1100MS, T#1700MS, T#1500MS, T#3500MS, T#2100MS, T#1700MS, T#1100MS, T#1700MS, T#2300MS, T#2400MS, T#1300MS, T#1700MS, T#1100MS, T#1700MS, T#1500MS, T#2400MS, T#2100MS, T#1700MS, T#1100MS, T#1700MS, T#2300MS];
    WD_RETRIEVE : ARRAY[1..12, 1..12] OF TIME := [T#6000MS, T#2100MS, T#1700MS, T#1100MS, T#1700MS, T#1900MS, T#6000MS, T#2100MS, T#1700MS, T#1100MS, T#1700MS, T#2300MS, T#4800MS, T#2100MS, T#1700MS, T#1100MS, T#1700MS, T#1900MS, T#4800MS, T#2100MS, T#1700MS, T#1100MS, T#1700MS, T#2300MS, T#3500MS, T#2100MS, T#1700MS, T#1100MS, T#1700MS, T#1900MS, T#3500MS, T#2100MS, T#1700MS, T#1100MS, T#1700MS, T#2300MS, T#2400MS, T#2100MS, T#1700MS, T#1100MS, T#1700MS, T#1900MS, T#2400MS, T#2100MS, T#1700MS, T#1100MS, T#1700MS, T#2300MS, T#6000MS, T#1100MS, T#1700MS, T#1100MS, T#1700MS, T#1100MS, T#6000MS, T#2100MS, T#1700MS, T#1100MS, T#1700MS, T#2300MS, T#4800MS, T#1100MS, T#1700MS, T#1100MS, T#1700MS, T#1100MS, T#4800MS, T#2100MS, T#1700MS, T#1100MS, T#1700MS, T#2300MS, T#3500MS, T#1100MS, T#1700MS, T#1100MS, T#1700MS, T#1100MS, T#3500MS, T#2100MS, T#1700MS, T#1100MS, T#1700MS, T#2300MS, T#2400MS, T#1100MS, T#1700MS, T#1100MS, T#1700MS, T#1100MS, T#2400MS, T#2100MS, T#1700MS, T#1100MS, T#1700MS, T#2300MS, T#6000MS, T#1300MS, T#1700MS, T#1100MS, T#1700MS, T#1500MS, T#6000MS, T#2100MS, T#1700MS, T#1100MS, T#1700MS, T#2300MS, T#4800MS, T#1300MS, T#1700MS, T#1100MS, T#1700MS, T#1500MS, T#4800MS, T#2100MS, T#1700MS, T#1100MS, T#1700MS, T#2300MS, T#3500MS, T#1300MS, T#1700MS, T#1100MS, T#1700MS, T#1500MS, T#3500MS, T#2100MS, T#1700MS, T#1100MS, T#1700MS, T#2300MS, T#2400MS, T#1300MS, T#1700MS, T#1100MS, T#1700MS, T#1500MS, T#2400MS, T#2100MS, T#1700MS, T#1100MS, T#1700MS, T#2300MS];
END_VAR

(* every scan: outputs off unless the active state sets them; Done is a pulse *)
Q3 := FALSE; Q4 := FALSE; Q5 := FALSE; Q6 := FALSE; Q7 := FALSE; Q8 := FALSE; Done := FALSE;
IF NOT Enable AND Sn <> 900 THEN Sn := 900; END_IF;
Wd(IN := (Sn = Prev) AND (WdTime > T#0MS), PT := WdTime);
Tm(IN := (Sn = Prev), PT := T#1H);
Prev := Sn;
IF Wd.Q THEN Alarm := Sn; Sn := 910; END_IF;

CASE Sn OF
  0: (* INIT: power-up, all outputs off *)
      WdTime := T#0MS; IF Enable THEN Sn := 10; END_IF;
  10: (* H:fork: Ausleger back to its rear stop *)
      WdTime := T#1700MS;
      Q8 := TRUE;
      IF I6 THEN Sn := 11; END_IF;
  11: (* H:lift: lift to the reference switch (direction ASSUMED: down) *)
      WdTime := T#3300MS;
      Q5 := TRUE;
      IF I4 THEN Sn := 12; END_IF;
  12: (* H:travel: travel to the reference switch (direction ASSUMED: to the belt) *)
      WdTime := T#6000MS;
      Q4 := TRUE;
      IF I1 THEN Sn := 13; END_IF;
  13: (* H:transit: lift to transit height (the pose every job starts from) *)
      WdTime := T#3100MS;
      CASE Drive(PosLift, 260.0, 0.375) OF -1: Q5 := TRUE; 1: Q6 := TRUE; END_CASE;
      IF ABS(PosLift - 260.0) <= 1.0 THEN Sn := 100; END_IF;
  100: (* READY: homed, waiting for a job *)
      WdTime := T#0MS; Ready := TRUE; Busy := FALSE;
      IF Cmd <> 0 THEN Job := Cmd; B1 := Arg1; Busy := TRUE; Ready := FALSE;
          CASE Cmd OF 11: Sn := 1000; 13: Sn := 2000; 14: Sn := 3000; 15: Sn := 4000; ELSE Sn := 910; Alarm := -Cmd; END_CASE;
      END_IF;
  1000: (* store_retrieve.01 lift->80: lift to 80 *)
      WdTime := T#2300MS;
      CASE Drive(PosLift, TG_STORE_RETRIEVE_LIFT[B1, 1], 0.375) OF -1: Q5 := TRUE; 1: Q6 := TRUE; END_CASE;
      IF ABS(PosLift - TG_STORE_RETRIEVE_LIFT[B1, 1]) <= 1.0 THEN Sn := 1001; END_IF;
  1001: (* store_retrieve.02 fork->out: Ausleger out to its front stop *)
      WdTime := T#1700MS;
      Q7 := TRUE;
      IF I5 THEN Sn := 1002; END_IF;
  1002: (* store_retrieve.03 lift->100: lift to 100 *)
      WdTime := T#1100MS;
      CASE Drive(PosLift, TG_STORE_RETRIEVE_LIFT[B1, 3], 0.375) OF -1: Q5 := TRUE; 1: Q6 := TRUE; END_CASE;
      IF ABS(PosLift - TG_STORE_RETRIEVE_LIFT[B1, 3]) <= 1.0 THEN Sn := 1003; END_IF;
  1003: (* store_retrieve.04 fork->back: Ausleger back to its rear stop *)
      WdTime := T#1700MS;
      Q8 := TRUE;
      IF I6 THEN Sn := 1004; END_IF;
  1004: (* store_retrieve.05 lift->tr: lift to transit *)
      WdTime := T#2100MS;
      CASE Drive(PosLift, TG_STORE_RETRIEVE_LIFT[B1, 5], 0.375) OF -1: Q5 := TRUE; 1: Q6 := TRUE; END_CASE;
      IF ABS(PosLift - TG_STORE_RETRIEVE_LIFT[B1, 5]) <= 1.0 THEN Sn := 1005; END_IF;
  1005: (* store_retrieve.06 travel->col: travel to the slot column *)
      WdTime := WD_STORE_RETRIEVE[B1, 6];
      CASE Drive(PosTravel, TG_STORE_RETRIEVE_TRAVEL[B1, 6], 0.375) OF -1: Q3 := TRUE; 1: Q4 := TRUE; END_CASE;
      IF ABS(PosTravel - TG_STORE_RETRIEVE_TRAVEL[B1, 6]) <= 1.0 THEN Sn := 1006; END_IF;
  1006: (* store_retrieve.07 lift->row: lift to row *)
      WdTime := WD_STORE_RETRIEVE[B1, 7];
      CASE Drive(PosLift, TG_STORE_RETRIEVE_LIFT[B1, 7], 0.375) OF -1: Q5 := TRUE; 1: Q6 := TRUE; END_CASE;
      IF ABS(PosLift - TG_STORE_RETRIEVE_LIFT[B1, 7]) <= 1.0 THEN Sn := 1007; END_IF;
  1007: (* store_retrieve.08 fork->out: Ausleger out to its front stop *)
      WdTime := T#1700MS;
      Q7 := TRUE;
      IF I5 THEN Sn := 1008; END_IF;
  1008: (* store_retrieve.09 lift->row-20: lift to row-20 *)
      WdTime := T#1100MS;
      CASE Drive(PosLift, TG_STORE_RETRIEVE_LIFT[B1, 9], 0.375) OF -1: Q5 := TRUE; 1: Q6 := TRUE; END_CASE;
      IF ABS(PosLift - TG_STORE_RETRIEVE_LIFT[B1, 9]) <= 1.0 THEN Sn := 1009; END_IF;
  1009: (* store_retrieve.10 fork->back: Ausleger back to its rear stop *)
      WdTime := T#1700MS;
      Q8 := TRUE;
      IF I6 THEN Sn := 1010; END_IF;
  1010: (* store_retrieve.11 lift->tr: lift to transit *)
      WdTime := WD_STORE_RETRIEVE[B1, 11];
      CASE Drive(PosLift, TG_STORE_RETRIEVE_LIFT[B1, 11], 0.375) OF -1: Q5 := TRUE; 1: Q6 := TRUE; END_CASE;
      IF ABS(PosLift - TG_STORE_RETRIEVE_LIFT[B1, 11]) <= 1.0 THEN Sn := 1011; END_IF;
  1011: (* store_retrieve.12 travel->col: travel to the next slot's column *)
      WdTime := WD_STORE_RETRIEVE[B1, 12];
      CASE Drive(PosTravel, TG_STORE_RETRIEVE_TRAVEL[B1, 12], 0.375) OF -1: Q3 := TRUE; 1: Q4 := TRUE; END_CASE;
      IF ABS(PosTravel - TG_STORE_RETRIEVE_TRAVEL[B1, 12]) <= 1.0 THEN Sn := 1012; END_IF;
  1012: (* store_retrieve.13 lift->row-20: lift to row-20 *)
      WdTime := WD_STORE_RETRIEVE[B1, 13];
      CASE Drive(PosLift, TG_STORE_RETRIEVE_LIFT[B1, 13], 0.375) OF -1: Q5 := TRUE; 1: Q6 := TRUE; END_CASE;
      IF ABS(PosLift - TG_STORE_RETRIEVE_LIFT[B1, 13]) <= 1.0 THEN Sn := 1013; END_IF;
  1013: (* store_retrieve.14 fork->out: Ausleger out to its front stop *)
      WdTime := T#1700MS;
      Q7 := TRUE;
      IF I5 THEN Sn := 1014; END_IF;
  1014: (* store_retrieve.15 lift->row: lift to row *)
      WdTime := T#1100MS;
      CASE Drive(PosLift, TG_STORE_RETRIEVE_LIFT[B1, 15], 0.375) OF -1: Q5 := TRUE; 1: Q6 := TRUE; END_CASE;
      IF ABS(PosLift - TG_STORE_RETRIEVE_LIFT[B1, 15]) <= 1.0 THEN Sn := 1015; END_IF;
  1015: (* store_retrieve.16 fork->back: Ausleger back to its rear stop *)
      WdTime := T#1700MS;
      Q8 := TRUE;
      IF I6 THEN Sn := 1016; END_IF;
  1016: (* store_retrieve.17 lift->tr: lift to transit *)
      WdTime := WD_STORE_RETRIEVE[B1, 17];
      CASE Drive(PosLift, TG_STORE_RETRIEVE_LIFT[B1, 17], 0.375) OF -1: Q5 := TRUE; 1: Q6 := TRUE; END_CASE;
      IF ABS(PosLift - TG_STORE_RETRIEVE_LIFT[B1, 17]) <= 1.0 THEN Sn := 1017; END_IF;
  1017: (* store_retrieve.18 travel->cv: travel to the conveyor *)
      WdTime := WD_STORE_RETRIEVE[B1, 18];
      CASE Drive(PosTravel, TG_STORE_RETRIEVE_TRAVEL[B1, 18], 0.375) OF -1: Q3 := TRUE; 1: Q4 := TRUE; END_CASE;
      IF ABS(PosTravel - TG_STORE_RETRIEVE_TRAVEL[B1, 18]) <= 1.0 THEN Sn := 1018; END_IF;
  1018: (* store_retrieve.19 lift->100: lift to 100 *)
      WdTime := T#2100MS;
      CASE Drive(PosLift, TG_STORE_RETRIEVE_LIFT[B1, 19], 0.375) OF -1: Q5 := TRUE; 1: Q6 := TRUE; END_CASE;
      IF ABS(PosLift - TG_STORE_RETRIEVE_LIFT[B1, 19]) <= 1.0 THEN Sn := 1019; END_IF;
  1019: (* store_retrieve.20 fork->out: Ausleger out to its front stop *)
      WdTime := T#1700MS;
      Q7 := TRUE;
      IF I5 THEN Sn := 1020; END_IF;
  1020: (* store_retrieve.21 lift->80: lift to 80 *)
      WdTime := T#1100MS;
      CASE Drive(PosLift, TG_STORE_RETRIEVE_LIFT[B1, 21], 0.375) OF -1: Q5 := TRUE; 1: Q6 := TRUE; END_CASE;
      IF ABS(PosLift - TG_STORE_RETRIEVE_LIFT[B1, 21]) <= 1.0 THEN Sn := 1021; END_IF;
  1021: (* store_retrieve.22 fork->back: Ausleger back to its rear stop *)
      WdTime := T#1700MS;
      Q8 := TRUE;
      IF I6 THEN Sn := 1022; END_IF;
  1022: (* store_retrieve.23 lift->tr: lift to transit *)
      WdTime := T#2300MS;
      CASE Drive(PosLift, TG_STORE_RETRIEVE_LIFT[B1, 23], 0.375) OF -1: Q5 := TRUE; 1: Q6 := TRUE; END_CASE;
      IF ABS(PosLift - TG_STORE_RETRIEVE_LIFT[B1, 23]) <= 1.0 THEN Done := TRUE; Busy := FALSE; Sn := 100; END_IF;
  2000: (* store.01 lift->80: lift to 80 *)
      WdTime := T#2300MS;
      CASE Drive(PosLift, TG_STORE_LIFT[B1, 1], 0.375) OF -1: Q5 := TRUE; 1: Q6 := TRUE; END_CASE;
      IF ABS(PosLift - TG_STORE_LIFT[B1, 1]) <= 1.0 THEN Sn := 2001; END_IF;
  2001: (* store.02 fork->out: Ausleger out to its front stop *)
      WdTime := T#1700MS;
      Q7 := TRUE;
      IF I5 THEN Sn := 2002; END_IF;
  2002: (* store.03 lift->100: lift to 100 *)
      WdTime := T#1100MS;
      CASE Drive(PosLift, TG_STORE_LIFT[B1, 3], 0.375) OF -1: Q5 := TRUE; 1: Q6 := TRUE; END_CASE;
      IF ABS(PosLift - TG_STORE_LIFT[B1, 3]) <= 1.0 THEN Sn := 2003; END_IF;
  2003: (* store.04 fork->back: Ausleger back to its rear stop *)
      WdTime := T#1700MS;
      Q8 := TRUE;
      IF I6 THEN Sn := 2004; END_IF;
  2004: (* store.05 lift->tr: lift to transit *)
      WdTime := T#2100MS;
      CASE Drive(PosLift, TG_STORE_LIFT[B1, 5], 0.375) OF -1: Q5 := TRUE; 1: Q6 := TRUE; END_CASE;
      IF ABS(PosLift - TG_STORE_LIFT[B1, 5]) <= 1.0 THEN Sn := 2005; END_IF;
  2005: (* store.06 travel->col: travel to the slot column *)
      WdTime := WD_STORE[B1, 6];
      CASE Drive(PosTravel, TG_STORE_TRAVEL[B1, 6], 0.375) OF -1: Q3 := TRUE; 1: Q4 := TRUE; END_CASE;
      IF ABS(PosTravel - TG_STORE_TRAVEL[B1, 6]) <= 1.0 THEN Sn := 2006; END_IF;
  2006: (* store.07 lift->row: lift to row *)
      WdTime := WD_STORE[B1, 7];
      CASE Drive(PosLift, TG_STORE_LIFT[B1, 7], 0.375) OF -1: Q5 := TRUE; 1: Q6 := TRUE; END_CASE;
      IF ABS(PosLift - TG_STORE_LIFT[B1, 7]) <= 1.0 THEN Sn := 2007; END_IF;
  2007: (* store.08 fork->out: Ausleger out to its front stop *)
      WdTime := T#1700MS;
      Q7 := TRUE;
      IF I5 THEN Sn := 2008; END_IF;
  2008: (* store.09 lift->row-20: lift to row-20 *)
      WdTime := T#1100MS;
      CASE Drive(PosLift, TG_STORE_LIFT[B1, 9], 0.375) OF -1: Q5 := TRUE; 1: Q6 := TRUE; END_CASE;
      IF ABS(PosLift - TG_STORE_LIFT[B1, 9]) <= 1.0 THEN Sn := 2009; END_IF;
  2009: (* store.10 fork->back: Ausleger back to its rear stop *)
      WdTime := T#1700MS;
      Q8 := TRUE;
      IF I6 THEN Sn := 2010; END_IF;
  2010: (* store.11 lift->tr: lift to transit *)
      WdTime := WD_STORE[B1, 11];
      CASE Drive(PosLift, TG_STORE_LIFT[B1, 11], 0.375) OF -1: Q5 := TRUE; 1: Q6 := TRUE; END_CASE;
      IF ABS(PosLift - TG_STORE_LIFT[B1, 11]) <= 1.0 THEN Sn := 2011; END_IF;
  2011: (* store.12 travel->cv: travel to the conveyor *)
      WdTime := WD_STORE[B1, 12];
      CASE Drive(PosTravel, TG_STORE_TRAVEL[B1, 12], 0.375) OF -1: Q3 := TRUE; 1: Q4 := TRUE; END_CASE;
      IF ABS(PosTravel - TG_STORE_TRAVEL[B1, 12]) <= 1.0 THEN Done := TRUE; Busy := FALSE; Sn := 100; END_IF;
  3000: (* fetch_empty.01 travel->col: travel to the slot column *)
      WdTime := WD_FETCH_EMPTY[B1, 1];
      CASE Drive(PosTravel, TG_FETCH_EMPTY_TRAVEL[B1, 1], 0.375) OF -1: Q3 := TRUE; 1: Q4 := TRUE; END_CASE;
      IF ABS(PosTravel - TG_FETCH_EMPTY_TRAVEL[B1, 1]) <= 1.0 THEN Sn := 3001; END_IF;
  3001: (* fetch_empty.02 lift->row-20: lift to row-20 *)
      WdTime := WD_FETCH_EMPTY[B1, 2];
      CASE Drive(PosLift, TG_FETCH_EMPTY_LIFT[B1, 2], 0.375) OF -1: Q5 := TRUE; 1: Q6 := TRUE; END_CASE;
      IF ABS(PosLift - TG_FETCH_EMPTY_LIFT[B1, 2]) <= 1.0 THEN Sn := 3002; END_IF;
  3002: (* fetch_empty.03 fork->out: Ausleger out to its front stop *)
      WdTime := T#1700MS;
      Q7 := TRUE;
      IF I5 THEN Sn := 3003; END_IF;
  3003: (* fetch_empty.04 lift->row: lift to row *)
      WdTime := T#1100MS;
      CASE Drive(PosLift, TG_FETCH_EMPTY_LIFT[B1, 4], 0.375) OF -1: Q5 := TRUE; 1: Q6 := TRUE; END_CASE;
      IF ABS(PosLift - TG_FETCH_EMPTY_LIFT[B1, 4]) <= 1.0 THEN Sn := 3004; END_IF;
  3004: (* fetch_empty.05 fork->back: Ausleger back to its rear stop *)
      WdTime := T#1700MS;
      Q8 := TRUE;
      IF I6 THEN Sn := 3005; END_IF;
  3005: (* fetch_empty.06 lift->tr: lift to transit *)
      WdTime := WD_FETCH_EMPTY[B1, 6];
      CASE Drive(PosLift, TG_FETCH_EMPTY_LIFT[B1, 6], 0.375) OF -1: Q5 := TRUE; 1: Q6 := TRUE; END_CASE;
      IF ABS(PosLift - TG_FETCH_EMPTY_LIFT[B1, 6]) <= 1.0 THEN Sn := 3006; END_IF;
  3006: (* fetch_empty.07 travel->cv: travel to the conveyor *)
      WdTime := WD_FETCH_EMPTY[B1, 7];
      CASE Drive(PosTravel, TG_FETCH_EMPTY_TRAVEL[B1, 7], 0.375) OF -1: Q3 := TRUE; 1: Q4 := TRUE; END_CASE;
      IF ABS(PosTravel - TG_FETCH_EMPTY_TRAVEL[B1, 7]) <= 1.0 THEN Sn := 3007; END_IF;
  3007: (* fetch_empty.08 lift->100: lift to 100 *)
      WdTime := T#2100MS;
      CASE Drive(PosLift, TG_FETCH_EMPTY_LIFT[B1, 8], 0.375) OF -1: Q5 := TRUE; 1: Q6 := TRUE; END_CASE;
      IF ABS(PosLift - TG_FETCH_EMPTY_LIFT[B1, 8]) <= 1.0 THEN Sn := 3008; END_IF;
  3008: (* fetch_empty.09 fork->out: Ausleger out to its front stop *)
      WdTime := T#1700MS;
      Q7 := TRUE;
      IF I5 THEN Sn := 3009; END_IF;
  3009: (* fetch_empty.10 lift->80: lift to 80 *)
      WdTime := T#1100MS;
      CASE Drive(PosLift, TG_FETCH_EMPTY_LIFT[B1, 10], 0.375) OF -1: Q5 := TRUE; 1: Q6 := TRUE; END_CASE;
      IF ABS(PosLift - TG_FETCH_EMPTY_LIFT[B1, 10]) <= 1.0 THEN Sn := 3010; END_IF;
  3010: (* fetch_empty.11 fork->back: Ausleger back to its rear stop *)
      WdTime := T#1700MS;
      Q8 := TRUE;
      IF I6 THEN Sn := 3011; END_IF;
  3011: (* fetch_empty.12 lift->tr: lift to transit *)
      WdTime := T#2300MS;
      CASE Drive(PosLift, TG_FETCH_EMPTY_LIFT[B1, 12], 0.375) OF -1: Q5 := TRUE; 1: Q6 := TRUE; END_CASE;
      IF ABS(PosLift - TG_FETCH_EMPTY_LIFT[B1, 12]) <= 1.0 THEN Done := TRUE; Busy := FALSE; Sn := 100; END_IF;
  4000: (* retrieve.01 travel->col: travel to the slot column *)
      WdTime := WD_RETRIEVE[B1, 1];
      CASE Drive(PosTravel, TG_RETRIEVE_TRAVEL[B1, 1], 0.375) OF -1: Q3 := TRUE; 1: Q4 := TRUE; END_CASE;
      IF ABS(PosTravel - TG_RETRIEVE_TRAVEL[B1, 1]) <= 1.0 THEN Sn := 4001; END_IF;
  4001: (* retrieve.02 lift->row-20: lift to row-20 *)
      WdTime := WD_RETRIEVE[B1, 2];
      CASE Drive(PosLift, TG_RETRIEVE_LIFT[B1, 2], 0.375) OF -1: Q5 := TRUE; 1: Q6 := TRUE; END_CASE;
      IF ABS(PosLift - TG_RETRIEVE_LIFT[B1, 2]) <= 1.0 THEN Sn := 4002; END_IF;
  4002: (* retrieve.03 fork->out: Ausleger out to its front stop *)
      WdTime := T#1700MS;
      Q7 := TRUE;
      IF I5 THEN Sn := 4003; END_IF;
  4003: (* retrieve.04 lift->row: lift to row *)
      WdTime := T#1100MS;
      CASE Drive(PosLift, TG_RETRIEVE_LIFT[B1, 4], 0.375) OF -1: Q5 := TRUE; 1: Q6 := TRUE; END_CASE;
      IF ABS(PosLift - TG_RETRIEVE_LIFT[B1, 4]) <= 1.0 THEN Sn := 4004; END_IF;
  4004: (* retrieve.05 fork->back: Ausleger back to its rear stop *)
      WdTime := T#1700MS;
      Q8 := TRUE;
      IF I6 THEN Sn := 4005; END_IF;
  4005: (* retrieve.06 lift->tr: lift to transit *)
      WdTime := WD_RETRIEVE[B1, 6];
      CASE Drive(PosLift, TG_RETRIEVE_LIFT[B1, 6], 0.375) OF -1: Q5 := TRUE; 1: Q6 := TRUE; END_CASE;
      IF ABS(PosLift - TG_RETRIEVE_LIFT[B1, 6]) <= 1.0 THEN Sn := 4006; END_IF;
  4006: (* retrieve.07 travel->cv: travel to the conveyor *)
      WdTime := WD_RETRIEVE[B1, 7];
      CASE Drive(PosTravel, TG_RETRIEVE_TRAVEL[B1, 7], 0.375) OF -1: Q3 := TRUE; 1: Q4 := TRUE; END_CASE;
      IF ABS(PosTravel - TG_RETRIEVE_TRAVEL[B1, 7]) <= 1.0 THEN Sn := 4007; END_IF;
  4007: (* retrieve.08 lift->100: lift to 100 *)
      WdTime := T#2100MS;
      CASE Drive(PosLift, TG_RETRIEVE_LIFT[B1, 8], 0.375) OF -1: Q5 := TRUE; 1: Q6 := TRUE; END_CASE;
      IF ABS(PosLift - TG_RETRIEVE_LIFT[B1, 8]) <= 1.0 THEN Sn := 4008; END_IF;
  4008: (* retrieve.09 fork->out: Ausleger out to its front stop *)
      WdTime := T#1700MS;
      Q7 := TRUE;
      IF I5 THEN Sn := 4009; END_IF;
  4009: (* retrieve.10 lift->80: lift to 80 *)
      WdTime := T#1100MS;
      CASE Drive(PosLift, TG_RETRIEVE_LIFT[B1, 10], 0.375) OF -1: Q5 := TRUE; 1: Q6 := TRUE; END_CASE;
      IF ABS(PosLift - TG_RETRIEVE_LIFT[B1, 10]) <= 1.0 THEN Sn := 4010; END_IF;
  4010: (* retrieve.11 fork->back: Ausleger back to its rear stop *)
      WdTime := T#1700MS;
      Q8 := TRUE;
      IF I6 THEN Sn := 4011; END_IF;
  4011: (* retrieve.12 lift->tr: lift to transit *)
      WdTime := T#2300MS;
      CASE Drive(PosLift, TG_RETRIEVE_LIFT[B1, 12], 0.375) OF -1: Q5 := TRUE; 1: Q6 := TRUE; END_CASE;
      IF ABS(PosLift - TG_RETRIEVE_LIFT[B1, 12]) <= 1.0 THEN Done := TRUE; Busy := FALSE; Sn := 100; END_IF;
  900: (* ESTOP: the safety relay dropped, outputs off *)
      WdTime := T#0MS; Busy := FALSE; Ready := FALSE; IF Reset AND Enable THEN Sn := 0; END_IF;
  910: (* FAULT: a step timed out, outputs off, alarm raised *)
      WdTime := T#0MS; Fault := TRUE; Busy := FALSE; Ready := FALSE;
      IF Ack AND Enable THEN Fault := FALSE; Sn := 10; END_IF;
END_CASE;
END_FUNCTION_BLOCK
